(* IEC 61131-3 sources: daoli-st-library/DL_Device (part 24) *)

(* ---- FB_DL_HumidifierWaterQual.st ---- *)
(*
  FB_DL_HumidifierWaterQual  —  加湿器水质电导率监视与排水联锁 / Humidifier water conductivity monitoring with drain interlock
  分类 Category : DL_Device
  码位 Code     : 16#03_2_04
  版本 Version  : 1.0.0
  溯源 Source   : 道莅自研 clean-room（电导率标定与排水联锁为通用水处理工程语义）
  功能 Function : 1) 电导率经标定换算（斜率/偏置）后按门限分级，超标触发排水周期；
                  2) 排水阀与补水阀互斥，同拍双开即判冲突并双双回安全位（关阀）；
                  3) 电导门限带迟滞防抖，越限解除有可到达路径；标定斜率非法（0/负）即拒算并置码。
  边界 Boundary : ① 标定参数非法（斜率 0 或负）拒算并置码；
                  ② 排水联锁与补水阀互斥（同拍双开判冲突回安全位）；
                  ③ 电导门限带迟滞防抖，越限解除有可到达路径；
                  ④ 输出三行同向：电导值 → 分级 → 排水阀。
  依赖 Depends  : FC_DL_LimitClassify（电导分级，每拍无条件调用）、FB_DL_TimeWindowCheck（排水维护时间窗，每拍无条件调用）

  码表 Error codes（本件子码步进 16#10，避让邻件码位）:
    16#0002_0304 故障级：电导率标定参数非法（斜率 <= 0 或非有限），拒算
    16#0002_0314 故障级：排水阀与补水阀同拍双开（互斥冲突），双双回安全位
    16#0002_0324 信息级：电导率越限已启动排水（不置 bError）
*)

TYPE E_DL_HwqPhase :
(
    eIdle    := 0,   // 空闲 / Idle
    eMonitor := 10,  // 电导监视 / Conductivity monitoring
    eDrain   := 20,  // 排水周期进行 / Drain cycle running
    eHold    := 30,  // 拒算保持 / Rejected, held
    eFault   := 90   // 故障锁定 / Fault locked
);
END_TYPE

FUNCTION_BLOCK FB_DL_HumidifierWaterQual
VAR_INPUT
    bEnable      : BOOL;                          // 总使能，FALSE 关阀回空闲 / Master enable
    bReset       : BOOL;                          // 复位，上升沿清故障与冲突锁存 / Reset
    fCondRawUScm : REAL;                          // 电导率原始值 [uS/cm]，域 0~2000 / Raw conductivity [uS/cm]
    fCalSlope    : REAL := 1.0;                   // 电导标定斜率 [uS/cm per 原始计数]，域 > 0 / Calibration slope
    fCalOffset   : REAL := 0.0;                   // 电导标定偏置 [uS/cm] / Calibration offset [uS/cm]
    fCondWarnUScm: REAL := 300.0;                 // 电导警告门限 [uS/cm]，域 > 0 / Conductivity warning limit
    fCondTripUScm: REAL := 600.0;                 // 电导排水门限 [uS/cm]，须 > 警告门限 / Drain trigger limit
    fCondHystUScm: REAL := 20.0;                  // 电导迟滞 [uS/cm]，域 >= 0 / Conductivity hysteresis
    tDrainTime   : TIME := T#30S;                 // 单次排水时长 [ms]，域 > 0 / Drain duration [ms]
    tDrainPeriod : TIME := T#10M;                 // 排水周期 [ms]，域 > 0 / Drain period [ms]
    uHourNow     : USINT := 0;                    // 当前时刻-时 [h]（注入，禁读 CPU 钟）/ Injected hour [h]
    uMinNow      : USINT := 0;                    // 当前时刻-分 [min]（注入）/ Injected minute [min]
    fEps         : REAL := 1.0E-6;                // 浮点判零容差 [1] / Floating zero tolerance
END_VAR
VAR_OUTPUT
    fCondUScm    : REAL;                          // 标定后电导率 [uS/cm] / Calibrated conductivity [uS/cm]
    bDrainValve  : BOOL;                          // 排水阀 [开关] / Drain valve
    bFillValve   : BOOL;                          // 补水阀 [开关] / Make-up fill valve
    bCondWarn    : BOOL;                          // 电导警告（保持型）/ Conductivity warning, held
    bInDrainWin  : BOOL;                          // 处于维护排水时间窗 / Inside maintenance drain window
    bValveConflict : BOOL;                        // 阀门互斥冲突标志 / Valve exclusion conflict flag
    bError       : BOOL;                          // 故障标志，与故障级码配对 / Fault flag paired with fault codes
    uErrorId     : UDINT;                         // 事件码，0 = 无事件 / Event code, 0 = none
    eStateOut    : E_DL_HwqPhase;                 // 状态机当前态，段尾单点映射 / Phase mapped at tail
END_VAR
VAR
    _eState      : E_DL_HwqPhase := E_DL_HwqPhase.eIdle;  // 内部状态 / Internal state
    rtrReset     : R_TRIG;                        // 复位沿 / Reset edge
    tonDrain     : TON;                           // 排水时长计时（自复位）/ Drain duration timer
    tonPeriod    : TON;                           // 排水周期节拍（自复位）/ Drain period tick
    fbWindow     : FB_DL_TimeWindowCheck;         // 排水维护时间窗实例（无条件调用）/ Drain time window
    bCalOk       : BOOL;                          // 标定参数合法 / Calibration valid
    bCfgOk       : BOOL;                          // 组态合法 / Configuration valid
    eBand        : E_DL_LimitBand;                // 电导分级结果 / Conductivity band
    aDayEn       : ARRAY[1..7] OF BOOL;           // 星期使能表（周一~周日）/ Weekday enable table
    nDay         : INT;                           // 星期填充下标 / Weekday fill index
    fCondCal     : REAL;                          // 标定后电导率暂存 [uS/cm] / Calibrated conductivity buffer
    bCondHigh    : BOOL;                          // 越排水门限标志 / Above drain threshold
    bDrainCmd    : BOOL;                          // 排水指令暂存 / Drain command buffer
    bFillCmd     : BOOL;                          // 补水指令暂存 / Fill command buffer
    uFault       : UDINT;                         // 锁存故障码 / Latched fault code
    uInfo        : UDINT;                         // 信息级码 / Information code
END_VAR
VAR CONSTANT
    DL_HWQ_CMAX  : REAL := 2000.0;                // 电导物理域上限 [uS/cm] / Conductivity domain high
END_VAR

(* === 段 0 · 实例刷新（无条件周期调用，自复位节拍）=== *)
rtrReset(CLK := bReset);                          // 每拍刷新复位沿
tonDrain(IN := (_eState = E_DL_HwqPhase.eDrain) AND (NOT tonDrain.Q), PT := tDrainTime);   // 自复位
tonPeriod(IN := NOT tonPeriod.Q, PT := tDrainPeriod);                                      // 周期心跳自复位
FOR nDay := 1 TO 7 DO
    aDayEn[nDay] := TRUE;                         // 维护排水窗与星期无关：全周使能
END_FOR
fbWindow(uHourNow := uHourNow,                    // 注入当前时
         uMinNow := uMinNow,                      // 注入当前分
         bEnableDay := TRUE,                      // 日窗使能
         aWeekdayEnable := aDayEn,                // 周一到周日全开（本地数组填充）
         uWeekdayNow := 1,                        // 星期注入（维护窗与星期无关）
         uHourOn := 0,                            // 窗开 00:00
         uMinOn := 0,                             // 窗开 0 分
         uHourOff := 23,                          // 窗关 23:00
         uMinOff := 59,                           // 窗关 59 分
         bReset := rtrReset.Q);                   // 复位沿清信息码
bInDrainWin := fbWindow.bInWindow;                // 时间窗输出

(* === 段 1 · 标定与组态闸 === *)
bCalOk := (fCalSlope > fEps) AND (fCalSlope = fCalSlope) AND (fCalOffset = fCalOffset);   // 斜率正域 + NaN 自反
bCfgOk := (fCondWarnUScm > fEps) AND (fCondTripUScm > fCondWarnUScm)
          AND (fCondHystUScm >= 0.0) AND (tDrainTime > T#0MS) AND (tDrainPeriod > T#0MS)
          AND (fCondWarnUScm = fCondWarnUScm) AND (fCondTripUScm = fCondTripUScm);   // 含 NaN 自反
IF NOT bCalOk THEN
    uFault := 16#0002_0304;                       // 故障级：标定参数非法，拒算
END_IF
IF NOT bCfgOk THEN
    uFault := 16#0002_0304;                       // 故障级：组态非法同码段（防无码可查）
END_IF
IF rtrReset.Q AND bCalOk AND bCfgOk THEN
    uFault := 16#0000;                            // 复位沿清锁存（复位路径可达）
    bValveConflict := FALSE;                      // 冲突标志同步复位
    bCondWarn := FALSE;                           // 警告标志同步复位
END_IF
uInfo := 16#0000;                                 // 信息码每拍清零
IF bCalOk AND (fCondRawUScm = fCondRawUScm) AND (fCondRawUScm >= 0.0)
   AND (fCondRawUScm <= DL_HWQ_CMAX) THEN
    fCondCal := fCondRawUScm * fCalSlope + fCalOffset;   // 标定换算
    IF fCondCal < 0.0 THEN
        fCondCal := 0.0;                          // 负电导截零（物理不可达）
    END_IF
    fCondUScm := fCondCal;                        // 电导值输出
ELSE
    fCondCal := 0.0;                              // 拒算：不出数值
END_IF

(* === 段 2 · 电导分级（函数每拍无条件调用）=== *)
eBand := FC_DL_LimitClassify(fVal := fCondCal,
                             fLowLimit := -1.0,               // 低低限：本件不使用（负值域）
                             fLowWarn := -0.5,                // 低警告限：本件不使用
                             fUpWarn := fCondWarnUScm,        // 高警告限
                             fUpLimit := fCondTripUScm);      // 高排水限
bCondHigh := (eBand = E_DL_LimitBand.eUpTripped);  // 到达排水级
IF eBand = E_DL_LimitBand.eUpWarn THEN
    bCondWarn := TRUE;                             // 警告级：置警告
END_IF

(* === 段 3 · 主状态机（ENUM + CASE，含 ELSE 兜底）=== *)
CASE _eState OF
E_DL_HwqPhase.eIdle :
    bDrainCmd := FALSE;                            // 空闲不排水
    bFillCmd := FALSE;                             // 空闲不补水
    IF (uFault <> 16#0000) AND (uFault <> 16#0002_0314) THEN
        _eState := E_DL_HwqPhase.eFault;           // 故障优先
    ELSIF bEnable AND (NOT bCalOk) THEN
        _eState := E_DL_HwqPhase.eHold;            // 标定非法：拒算保持
    ELSIF bEnable THEN
        _eState := E_DL_HwqPhase.eMonitor;         // 进入监视相
    END_IF

E_DL_HwqPhase.eMonitor :
    bFillCmd := NOT bDrainCmd;                     // 补水默认开（与排水互斥）
    IF bCondHigh THEN
        bCondWarn := TRUE;                         // 置位型：电导警告
        uInfo := 16#0002_0324;                     // 信息级：越限启动排水
        _eState := E_DL_HwqPhase.eDrain;           // 转排水相
    ELSIF (eBand = E_DL_LimitBand.eNormal) AND (fCondCal < (fCondWarnUScm - fCondHystUScm)) THEN
        bCondWarn := FALSE;                        // 迟滞带下方：解除警告（可到达的解除路径）
    END_IF
    IF (NOT bEnable) OR (NOT bCalOk) THEN
        _eState := E_DL_HwqPhase.eIdle;            // 失能/标定失效回空闲
    END_IF

E_DL_HwqPhase.eDrain :
    bDrainCmd := TRUE;                             // 排水阀开（驱动方向）
    bFillCmd := FALSE;                             // 补水阀关（互斥）
    IF tonDrain.Q THEN
        bDrainCmd := FALSE;                        // 排水时长到：关阀（本拍行为）
        IF bCondHigh THEN
            IF tonPeriod.Q THEN
                bFillCmd := TRUE;                  // 周期未到且仍超标：等待下一周期再排
            END_IF
            _eState := E_DL_HwqPhase.eMonitor;     // 回监视相，等下一周期
        ELSE
            _eState := E_DL_HwqPhase.eMonitor;     // 达标：回监视相
        END_IF
    END_IF

E_DL_HwqPhase.eHold :
    bDrainCmd := FALSE;                            // 拒算态关排水
    bFillCmd := FALSE;                             // 拒算态关补水
    IF bCalOk THEN
        _eState := E_DL_HwqPhase.eMonitor;         // 标定恢复：解除拒算（可到达的解除路径）
    END_IF

E_DL_HwqPhase.eFault :
    bDrainCmd := FALSE;                            // 故障态排水阀关（安全侧）
    bFillCmd := FALSE;                             // 故障态补水阀关
    IF uFault = 16#0000 THEN
        _eState := E_DL_HwqPhase.eIdle;            // 解锁回空闲
    END_IF

ELSE
    _eState := E_DL_HwqPhase.eFault;               // 非法状态拦截
    uFault := 16#0002_0304;                        // 故障级：相 ID 越界
    bDrainCmd := FALSE;                            // 安全侧关阀
    bFillCmd := FALSE;                             // 安全侧关阀
END_CASE

(* === 段 4 · 阀门互斥仲裁（同拍双开判冲突，双双回安全位）=== *)
IF bDrainCmd AND bFillCmd THEN
    bDrainCmd := FALSE;                            // 冲突：排水阀回安全位
    bFillCmd := FALSE;                             // 冲突：补水阀回安全位
    bValveConflict := TRUE;                        // 冲突标志置位
    uFault := 16#0002_0314;                        // 故障级：互斥冲突
ELSE
    bValveConflict := FALSE;                       // 无冲突：标志清零（非置位型）
END_IF
IF rtrReset.Q AND bValveConflict THEN
    uFault := 16#0000;                             // 冲突经复位解除（复位路径可达）
    bValveConflict := FALSE;                       // 标志同步清零
END_IF
IF NOT bEnable THEN
    bDrainCmd := FALSE;                            // 失能最高优先：排水关
    bFillCmd := FALSE;                             // 失能最高优先：补水关
END_IF

(* === 段 5 · 输出映射（三行同向：电导值 → 分级 → 排水阀）=== *)
bDrainValve := bDrainCmd;                          // 排水阀输出
bFillValve := bFillCmd;                            // 补水阀输出
bError := (uFault <> 16#0000);                     // 故障标志仅由故障级码置位（R45 配对）
IF bError THEN
    uErrorId := uFault;                            // 故障级优先上报
ELSE
    uErrorId := uInfo;                             // 否则上报信息级码
END_IF
eStateOut := _eState;                              // 输出枚举段尾单点映射（N2 规则）
END_FUNCTION_BLOCK

(* ---- FB_DL_HydraulicAccumPreChg.st ---- *)
(*
  ==================================================================
  组件名 Component  : FB_DL_HydraulicAccumPreChg
  分类   Category   : DL_Device
  复杂度 Complexity  : cx3
  版本   Version    : 1.0.1
  功能   Purpose    : 液压蓄能器氮气预充压力监视。把实测气囊压力按理想气体等温
                      折算到参考温度 20 摄氏度（pCorr = pGas · T0K / TK），再对额定
                      预充压力求偏差百分比；欠充 / 过充双态判据带迟滞防抖；油口
                      压力显著高于气囊侧判气囊失效疑点（eBladderSuspect）；传感器
                      非有限或压力 / 温度物理域越界判 eSensorBad。
  来源   Source     : t2-2-lbp
  溯源   Origin     : IEC 61131-3 标准语义的道莅防御性实现；理想气体等温折算与
                      蓄能器预充校验为公开热力学与液压语义，clean-room 自研实现，
                      未复制任何闭源代码行。
  平台   Platform   : 纯 IEC 61131-3（LREAL 运算，无私有库、无定时器实例）
  作者   Author     : 道莅代码库 · PLC 编程专家（R56）
  ------------------------------------------------------------------
  边界 Boundary     :
                      一 本件只做预充状态判级，不做充放气控制、不做泄放（属主边界）；
                      二 判据方向性（R146）：欠充与过充为同量纲双向异常，分派独立
                         成因成员（R190 归因唯一），互不合并；
                      三 迟滞口径：进入判据用全带宽，退出判据带宽收窄 fHystBar，
                         防边界抖动反复置清；
                      四 成因锁存解除路径 = bReset 上升沿（唯一路径，头注释声明，R188）；
                      五 无全局变量、无外部变量声明、无物理地址寻址。
  输出契约 Output contract:
                      fDevPct 为温度修正后偏差百分比（正 = 高于额定，负 = 低于额定）；
                      eFault 为锁存回放；bError 与故障级成因配对（R45）；
                      ePhaseBad 为非法相位兜底专用成员（R128）。
  修订记录 Revision  :
    2026-11-20  v1.0.0  R56 首版（批 2 · 序号 10）
    2026-11-21  v1.0.1  R57 返修：段 3 域闸补温度上界 150.0 摄氏度判 eSensorBad（阈值提为常量并注单位）
  ==================================================================
*)

TYPE E_DL_HapPhase :
(
    eIdle  := 0,  // 未使能：判级停摆 / disabled, the grading is idle
    eRun   := 10, // 运行：逐拍判级 / running, graded every scan
    eFault := 90  // 故障：成因锁存 / fault, the cause is latched
);
END_TYPE

TYPE E_DL_HapFault :
(
    eNone          := 0, // 无成因 / no cause
    eUnderCharge   := 1, // 预充不足（故障级，与 bError 配对）/ the precharge is under, fault grade paired with bError
    eOverCharge    := 2, // 预充过量（故障级，与 bError 配对）/ the precharge is over, fault grade paired with bError
    eBladderSuspect:= 3, // 油口压力显著高于气囊侧，气囊失效疑点（故障级，与 bError 配对）/ the oil side clearly exceeds the gas side, a bladder suspect, fault grade paired with bError
    eSensorBad     := 4, // 传感器非有限或物理域越界（故障级，与 bError 配对）/ a sensor is non finite or out of the physical domain, fault grade paired with bError
    ePhaseBad      := 5  // 非法相位兜底（故障级，与 bError 配对）/ illegal phase fallback, fault grade paired with bError
);
END_TYPE

FUNCTION_BLOCK FB_DL_HydraulicAccumPreChg
VAR_INPUT
    bEnable   : BOOL := TRUE;   // 使能，失能时判级停摆 [-] / enable, the grading stops when disabled
    bReset    : BOOL := FALSE;  // 复位上升沿清全部成因锁存 [-] / reset rising edge clears every cause latch
    pGas      : LREAL := 90.0;  // 气囊压力实测 [巴] / measured gas side pressure [bar]
    pOil      : LREAL := 0.0;   // 油口压力实测 [巴] / measured oil port pressure [bar]
    fTempC    : LREAL := 20.0;  // 气体温度实测 [摄氏度] / measured gas temperature [degree celsius]
    pNom      : LREAL := 90.0;  // 额定预充压力 [巴]，域 大于零 / rated precharge pressure [bar], domain above zero
    fUnderBar : LREAL := 9.0;   // 欠充判据带宽（低于额定的绝对量）[巴] / undercharge band below the rating [bar]
    fOverBar  : LREAL := 9.0;   // 过充判据带宽（高于额定的绝对量）[巴] / overcharge band above the rating [bar]
    fHystBar  : LREAL := 1.0;   // 迟滞带宽 [巴]，域 0..判据带宽 / hysteresis band [bar], inside the criterion band
    fBladMarg : LREAL := 20.0;  // 气囊疑点裕度（油口超出气囊侧百分比）[百分比] / bladder suspect margin over the gas side [percent]
END_VAR
VAR_OUTPUT
    fDevPct : LREAL := 0.0;  // 温度修正后预充偏差百分比 [百分比] / the corrected precharge deviation [percent]
    ePhase  : E_DL_HapPhase := E_DL_HapPhase.eIdle; // 相位出口 [枚举] / phase outlet [enum]
    eFault  : E_DL_HapFault := E_DL_HapFault.eNone; // 成因出口，锁存回放 [枚举] / cause outlet replayed from the latch [enum]
    bError  : BOOL := FALSE; // 故障锁存标志 [-] / fault latch flag
END_VAR
VAR
    rtReset  : R_TRIG; // 复位沿检测，段 0 无条件刷新 / reset edge, refreshed unconditionally in segment zero
    _ePhase  : E_DL_HapPhase := E_DL_HapPhase.eIdle; // 内部相位，CASE 唯一写入目标 / internal phase, the only CASE write target
    _eFaulC  : E_DL_HapFault := E_DL_HapFault.eNone; // 故障级成因，锁存至复位沿 / fault cause, latched until the reset edge
    _bFault  : BOOL := FALSE; // 故障锁存位 [-] / fault latch bit
    _bInit   : BOOL := FALSE; // 首扫初始化完成标志（R310）/ first scan initialisation flag
    _bInOk   : BOOL := FALSE; // 三个实数输入全部有限 [-] / all three real inputs are finite
    _bCfgOk  : BOOL := FALSE; // 组态参数域内 [-] / the configuration is inside the domain
    _fTK     : LREAL := 0.0;  // 气体绝对温度 [开尔文] / the absolute gas temperature [kelvin]
    _fPCorr  : LREAL := 0.0;  // 折算到参考温度的气囊压力 [巴] / the gas pressure corrected to the reference temperature [bar]
    _fDev    : LREAL := 0.0;  // 偏差绝对量 [巴] / the deviation magnitude [bar]
    _bUnder  : BOOL := FALSE; // 欠充迟滞锁存 [-] / the undercharge hysteresis latch
    _bOver   : BOOL := FALSE; // 过充迟滞锁存 [-] / the overcharge hysteresis latch
    _bBlad   : BOOL := FALSE; // 气囊疑点迟滞锁存 [-] / the bladder suspect hysteresis latch
    _bBad    : BOOL := FALSE; // 传感器无效锁存 [-] / the sensor bad latch
END_VAR
VAR CONSTANT
    DL_HAP_TEMP_HI : LREAL := 150.0; // 温度上界 [摄氏度]，超界判传感器无效（v1.0.1 返修）/ the temperature ceiling [degree celsius], beyond it the sensor is judged bad (v1.0.1 fix)
END_VAR

// 段 0｜沿检测无条件周期刷新（禁入分支）/ segment 0, unconditional refresh of the edge detector
rtReset(CLK := bReset); // 复位沿无条件刷新 / unconditional refresh of the reset edge

// 段 1｜首扫初始化（R310）/ segment 1, first scan initialisation
IF NOT _bInit THEN // 首扫一拍 / the very first scan
    _bInit := TRUE; // 置首扫完成标志 / raise the first scan flag
    _ePhase := E_DL_HapPhase.eRun; // 相位从运行起步（使能默认真）/ the phase starts in run
    _eFaulC := E_DL_HapFault.eNone; // 故障级成因清零 / clear the fault cause
    _bFault := FALSE; // 故障锁存清零 / clear the fault latch
END_IF

// 段 2｜复位沿作用域：清全部迟滞与锁存 / 迁相位（两项逐项声明）/ segment 2, reset edge scope declared item by item
IF rtReset.Q THEN // 复位沿 / the reset edge
    _bFault := FALSE; // 作用域一：清故障锁存 / scope one, clear the fault latch
    _eFaulC := E_DL_HapFault.eNone; // 作用域一：清故障级成因 / scope one, clear the fault cause
    _bUnder := FALSE; // 作用域一：清欠充迟滞 / scope one, clear the undercharge latch
    _bOver := FALSE; // 作用域一：清过充迟滞 / scope one, clear the overcharge latch
    _bBlad := FALSE; // 作用域一：清气囊疑点迟滞 / scope one, clear the bladder latch
    _bBad := FALSE; // 作用域一：清传感器无效锁存 / scope one, clear the sensor bad latch
    _ePhase := E_DL_HapPhase.eRun; // 作用域二：迁回运行相 / scope two, migrate back to run
END_IF

// 段 3｜组态与输入域闸（R151 全覆盖）/ segment 3, the configuration and input domain gates
_bInOk := (pGas = pGas) AND ((pGas - pGas) = (pGas - pGas)) AND (pOil = pOil) AND ((pOil - pOil) = (pOil - pOil)) AND (fTempC = fTempC) AND ((fTempC - fTempC) = (fTempC - fTempC)); // 三输入有限性 / finiteness of the three inputs
_bCfgOk := (pNom > 0.0) AND (pNom = pNom) AND (fUnderBar >= 0.0) AND (fUnderBar = fUnderBar) AND (fOverBar >= 0.0) AND (fOverBar = fOverBar) AND (fHystBar >= 0.0) AND (fHystBar <= fUnderBar) AND (fHystBar <= fOverBar) AND (fBladMarg > 0.0) AND (fBladMarg = fBladMarg); // 组态参数域判定 / the configuration domain verdict
IF (NOT _bInOk) OR (pGas < 0.0) OR (pOil < 0.0) OR (fTempC < -270.0) OR (fTempC > DL_HAP_TEMP_HI) OR (NOT _bCfgOk) THEN // 输入非有限、物理域越界（含 v1.0.1 温度上界）或组态非法 / a non finite input, a physical domain violation (with the v1.0.1 temperature ceiling) or an illegal configuration
    IF NOT _bBad THEN // 未锁存才置（防同拍抹除）/ set only while unlatched
        _bBad := TRUE; // 置传感器无效锁存 / raise the sensor bad latch
    END_IF
END_IF

// 段 4｜相位机：ENUM + CASE，含 ELSE 非法相位兜底（R128）/ segment 4, the phase machine with an ELSE fallback
CASE _ePhase OF
E_DL_HapPhase.eIdle: // 未使能相 / the disabled phase
    IF bEnable AND (NOT _bFault) THEN // 使能且无故障 / enabled and unfaulted
        _ePhase := E_DL_HapPhase.eRun; // 迁运行相 / migrate to run
    END_IF

E_DL_HapPhase.eRun: // 运行相：逐拍判级 / the run phase, graded every scan
    IF NOT bEnable THEN // 失能 / disabled
        _ePhase := E_DL_HapPhase.eIdle; // 迁未使能相 / migrate to idle
    ELSIF _bBad THEN // 传感器无效锁存优先 / the sensor bad latch takes priority
        _bFault := TRUE; // 置故障锁存 / raise the fault latch
        _eFaulC := E_DL_HapFault.eSensorBad; // 故障级成因（R45 配对 bError）/ the fault cause paired with bError
        _ePhase := E_DL_HapPhase.eFault; // 迁故障相 / migrate to the fault phase
    ELSE // 正常判级 / the normal grading
        _fTK := fTempC + 273.15; // 摄氏度转开尔文 / celsius to kelvin
        IF _fTK < 1.0 THEN // 绝对温度趋零防御（等温折算除子域闸）/ the absolute temperature guard for the divisor
            _fTK := 1.0; // 钳到下限 / clamp to the floor
        END_IF
        _fPCorr := pGas * (293.15 / _fTK); // 等温折算到 20 摄氏度参考（除子为绝对温度已证超阈）/ the isothermal correction to the twenty degree reference
        IF pNom > 0.0 THEN // 额定压力已证大于零（组态闸）/ the rating is proven positive by the gate
            fDevPct := (_fPCorr - pNom) / pNom * 100.0; // 偏差百分比 / the deviation percentage
        ELSE // 组态非法兜底（防御性保留）/ the illegal configuration fallback
            fDevPct := 0.0; // 偏差记零 / the deviation is zeroed
        END_IF
        _fDev := _fPCorr - pNom; // 偏差绝对量（带符号）/ the signed deviation
        IF _fDev < -fUnderBar THEN // 欠充进入判据 / the undercharge entry criterion
            _bUnder := TRUE; // 置欠充迟滞锁存 / raise the undercharge latch
        ELSIF _fDev > -fUnderBar + fHystBar THEN // 欠充退出判据（迟滞收窄）/ the undercharge exit criterion with the narrowed band
            _bUnder := FALSE; // 清欠充迟滞 / clear the undercharge latch
        END_IF
        IF _fDev > fOverBar THEN // 过充进入判据 / the overcharge entry criterion
            _bOver := TRUE; // 置过充迟滞锁存 / raise the overcharge latch
        ELSIF _fDev < fOverBar - fHystBar THEN // 过充退出判据（迟滞收窄）/ the overcharge exit criterion with the narrowed band
            _bOver := FALSE; // 清过充迟滞 / clear the overcharge latch
        END_IF
        IF pOil > _fPCorr * (1.0 + fBladMarg / 100.0) THEN // 油口显著高于气囊侧 / the oil side clearly exceeds the gas side
            _bBlad := TRUE; // 置气囊疑点迟滞锁存 / raise the bladder latch
        ELSIF pOil < _fPCorr * (1.0 + fBladMarg / 200.0) THEN // 气囊疑点退出判据（半带迟滞）/ the bladder exit criterion with a half band
            _bBlad := FALSE; // 清气囊疑点迟滞 / clear the bladder latch
        END_IF
        IF _bBlad THEN // 气囊疑点优先级最高（结构性失效）/ the bladder suspect has the highest priority, a structural failure
            _bFault := TRUE; // 置故障锁存 / raise the fault latch
            _eFaulC := E_DL_HapFault.eBladderSuspect; // 故障级成因（R45 配对 bError）/ the fault cause paired with bError
            _ePhase := E_DL_HapPhase.eFault; // 迁故障相 / migrate to the fault phase
        ELSIF _bOver THEN // 过充次优先 / the overcharge takes the next priority
            _bFault := TRUE; // 置故障锁存 / raise the fault latch
            _eFaulC := E_DL_HapFault.eOverCharge; // 故障级成因（R45 配对 bError）/ the fault cause paired with bError
            _ePhase := E_DL_HapPhase.eFault; // 迁故障相 / migrate to the fault phase
        ELSIF _bUnder THEN // 欠充再次优先 / the undercharge follows
            _bFault := TRUE; // 置故障锁存 / raise the fault latch
            _eFaulC := E_DL_HapFault.eUnderCharge; // 故障级成因（R45 配对 bError）/ the fault cause paired with bError
            _ePhase := E_DL_HapPhase.eFault; // 迁故障相 / migrate to the fault phase
        END_IF
    END_IF

E_DL_HapPhase.eFault: // 故障相：成因锁存，等待复位沿；偏差出口冻结保持末值（R191 显式声明）/ the fault phase, the cause is latched, the deviation outlet holds frozen

ELSE // 非法相位兜底（R128）/ the illegal phase fallback
    _bFault := TRUE; // 置故障锁存 / raise the fault latch
    _eFaulC := E_DL_HapFault.ePhaseBad; // 故障级成因（R45 配对 bError）/ the fault cause paired with bError
    _ePhase := E_DL_HapPhase.eFault; // 迁故障相 / migrate to the fault phase
END_CASE

// 段 5｜统一出口 / segment 5, the unified outlet
IF _bFault THEN // 故障锁存优先 / the fault latch takes priority
    eFault := _eFaulC; // 故障级成因锁存回放（不按当下输入重推断，R152）/ the fault cause replayed from the latch
ELSE
    eFault := E_DL_HapFault.eNone; // 无锁存即无成因 / no latch, no cause
END_IF
ePhase := _ePhase; // 相位出口单点映射 / single point phase outlet mapping
bError := _bFault; // 故障标志与锁存位同源 / the fault flag shares the latch source
END_FUNCTION_BLOCK

(* ---- FB_DL_HydroPressRampSeq.st ---- *)
(*
  ============================================================
  组件名 : FB_DL_HydroPressRampSeq
  分类   : DL_Device
  功能   : 液压建压斜坡顺序控制，建压升压保压泄压按斜率给定并含超时保护
  开源溯源 : internal-design（本轮无外部代码逐行引用）
             参考语义 : 无外部参考
  复杂度 : C2
  版本   : 1.0.0
  ============================================================
  配比约束 : tonRamp 与 tonHold 共用 tHoldTimeout 作为监视窗（升压窗与保压窗各一实例，
             两者互不累计）；tReleaseTimeout 单独覆盖泄压相。默认值须全部大于零。
  降级语义 : 实测压力非有限时冻结斜坡并保持上一有限设定输出，bPressOk 置假，不置故障码。
  故障码   : 1 保压超时 / 2 升压超时 / 3 泄压超时。码 3 不可由 1 与 2 观测——1 与 2 只在
             升压相与保压相置位，泄压相进入故障时码必为 0，故单开 3 以区分成因。
             复位唯一路径：bBuildCmd 或 bReleaseCmd 上升沿。
  ============================================================
*)

TYPE E_DL_HydroRampState :
(
    eIdle     := 0, // 待机，设定保持在零 idle with the set point at zero
    eRampUp   := 1, // 升压相，按斜率逼近目标 pressure ramp up towards the target
    eHold     := 2, // 保压相，设定保持目标 pressure hold at the target
    eRampDown := 3, // 泄压相，按斜率降到零 pressure ramp down to zero
    eFault    := 4  // 故障锁存相 latched fault phase
);
END_TYPE

FUNCTION_BLOCK FB_DL_HydroPressRampSeq
VAR_INPUT
    bBuildCmd      : BOOL; // 建压命令 pressure build command
    bReleaseCmd    : BOOL; // 泄压命令 pressure release command
    rPressAct      : REAL; // 实测压力 [bar] actual pressure [bar]
    rPressTarget   : REAL; // 目标压力 [bar] target pressure [bar]
    rRampBarPerS   : REAL; // 升压斜率 [bar/s] ramp rate [bar per second]
    rHoldBand      : REAL; // 保压允差带 [bar] hold band [bar]
    tHoldTimeout   : TIME; // 保压与升压监视窗 [ms] hold and ramp watchdog window
    tReleaseTimeout: TIME; // 泄压监视窗 [ms] release watchdog window
END_VAR
VAR_OUTPUT
    rPressSp   : REAL; // 压力设定输出 [bar] pressure set point [bar]
    eState     : E_DL_HydroRampState; // 当前状态 current state
    bPressOk   : BOOL; // 保压到位标志 pressure reached flag
    nFaultCode : INT; // 故障码 0无 1保压超时 2升压超时 3泄压超时 [码] fault code [code]
END_VAR
VAR
    _eState  : E_DL_HydroRampState := E_DL_HydroRampState.eIdle; // 内部状态 internal state
    _rSp     : REAL := 0.0; // 斜坡积分设定量 [bar] ramped set point [bar]
    _nFault  : INT := 0; // 故障码锁存内部量 latched fault code
    _bFin    : BOOL := FALSE; // 实数输入有限性判定 finiteness verdict of the real inputs
    _rBand   : REAL := 0.0; // 钳位后的允差带 [bar] clamped hold band [bar]
    tonTick  : TON; // 一秒节拍计时 one second tick timer
    tonHold  : TON; // 保压超时计时 hold timeout timer
    tonRamp  : TON; // 升压超时计时 ramp timeout timer
    tonRelease : TON; // 泄压超时计时 release timeout timer
    rtBuild  : R_TRIG; // 建压命令上升沿 build command rising edge
    rtRelease: R_TRIG; // 泄压命令上升沿 release command rising edge
END_VAR

// 段 0｜定时器与沿实例无条件周期刷新 unconditional cyclic refresh of timers and edges
tonTick(IN := NOT tonTick.Q, PT := T#1S); // 一秒自复位节拍 one second self reset tick
tonHold(IN := (_eState = E_DL_HydroRampState.eHold) AND (_nFault = 0), PT := tHoldTimeout); // 保压超时 hold timeout
tonRamp(IN := (_eState = E_DL_HydroRampState.eRampUp) AND (_nFault = 0), PT := tHoldTimeout); // 升压超时 ramp timeout
tonRelease(IN := (_eState = E_DL_HydroRampState.eRampDown) AND (_nFault = 0), PT := tReleaseTimeout); // 泄压超时 release timeout
rtBuild(CLK := bBuildCmd); // 建压沿刷新 refresh the build edge
rtRelease(CLK := bReleaseCmd); // 泄压沿刷新 refresh the release edge
// 段 1｜出口预置与输入整形 preset the outputs and reshape the inputs
bPressOk := FALSE; // 到位标志每拍先假 the reached flag is false each scan first
_rBand := rHoldBand; // 取入参允差带 take the hold band input
IF _rBand < 0.0 THEN
    _rBand := ABS(_rBand); // 负允差带取幅值 a negative band becomes its magnitude
END_IF
_bFin := (rPressAct = rPressAct) AND (rPressTarget = rPressTarget) AND (rRampBarPerS = rRampBarPerS) AND (rHoldBand = rHoldBand); // 四输入自反判定 self comparison of the four inputs
IF NOT _bFin THEN
    rPressSp := _rSp; // 冻结斜坡并输出上一有限设定 freeze the ramp and emit the last finite set point
    eState := _eState; // 状态出口按锁存量 map the state
    nFaultCode := _nFault; // 故障码出口按锁存量 map the fault code
    RETURN; // 非有限测量不迁相，早退 the non finite reading changes no phase
END_IF
// 段 2｜主状态机 main state machine
CASE _eState OF
E_DL_HydroRampState.eIdle: // 待机相 idle phase
    _rSp := 0.0; // 待机设定归零 the set point returns to zero
    IF rtBuild.Q AND (NOT bReleaseCmd) AND (rPressTarget > 0.0) AND (rRampBarPerS > 0.0) THEN
        _eState := E_DL_HydroRampState.eRampUp; // 组态合法才迁升压相 migrate only when the configuration is legal
    END_IF
E_DL_HydroRampState.eRampUp: // 升压相 ramp up phase
    IF tonTick.Q THEN
        _rSp := LIMIT(0.0, _rSp + rRampBarPerS, rPressTarget); // 每满一秒按斜率推进 advance one ramp step per full second
    END_IF
    IF (rPressAct >= (rPressTarget - _rBand)) AND (ABS(_rSp - rPressTarget) < 1.0E-3) THEN
        _eState := E_DL_HydroRampState.eHold; // 设定到位且反馈入带则迁保压 both the set point and the feedback are in place
    ELSIF tonRamp.Q THEN
        _nFault := 2; // 升压超时故障码 ramp timeout fault code
        _eState := E_DL_HydroRampState.eFault; // 迁故障相 migrate to the fault phase
    END_IF
E_DL_HydroRampState.eHold: // 保压相 hold phase
    _rSp := rPressTarget; // 设定保持目标 the set point holds the target
    IF ABS(rPressAct - rPressTarget) <= _rBand THEN
        bPressOk := TRUE; // 反馈在允差带内 the feedback sits inside the band
    END_IF
    IF rtRelease.Q OR bReleaseCmd THEN
        _eState := E_DL_HydroRampState.eRampDown; // 泄压命令优先于超时 the release command outranks the timeout
    ELSIF tonHold.Q THEN
        _nFault := 1; // 保压超时故障码 hold timeout fault code
        _eState := E_DL_HydroRampState.eFault; // 迁故障相 migrate to the fault phase
    END_IF
E_DL_HydroRampState.eRampDown: // 泄压相 ramp down phase
    IF tonTick.Q THEN
        _rSp := LIMIT(0.0, _rSp - rRampBarPerS, rPressTarget); // 每满一秒按斜率回落 fall one ramp step per full second
    END_IF
    IF (rPressAct < 0.5) AND (_rSp < 1.0E-3) THEN
        _rSp := 0.0; // 设定归零 the set point lands at zero
        _eState := E_DL_HydroRampState.eIdle; // 回待机 return to idle
    ELSIF tonRelease.Q THEN
        _nFault := 3; // 泄压超时故障码 release timeout fault code
        _eState := E_DL_HydroRampState.eFault; // 迁故障相 migrate to the fault phase
    END_IF
E_DL_HydroRampState.eFault: // 故障锁存相 latched fault phase
    IF rtBuild.Q OR rtRelease.Q THEN
        _nFault := 0; // 复位清故障码 the reset edge clears the fault code
        _rSp := 0.0; // 复位设定归零 the reset edge clears the set point
        _eState := E_DL_HydroRampState.eIdle; // 复位回待机 the reset edge returns to idle
    END_IF
ELSE // 非法状态枚举兜底 the illegal state fallback
    _eState := E_DL_HydroRampState.eIdle; // 非法状态回落待机 an illegal state falls back to idle
END_CASE
// 段 3｜统一出口映射 the unified exit mapping
rPressSp := _rSp; // 设定出口 map the set point
eState := _eState; // 状态出口 map the state
nFaultCode := _nFault; // 故障码出口 map the fault code
END_FUNCTION_BLOCK

(* ---- FB_DL_InductionHardeningScanCtrl.st ---- *)
(*
  Component : FB_DL_InductionHardeningScanCtrl
  Category  : DL_Device
  Type      : FB
  Complexity: C2
  VERSION   : v1.0.0
  功能      : 感应淬火扫描时序控制：ENUM 七态状态机（Idle/Heat/Scan/Spray/Cool/Done/Fault），扫描功率随速度联动，喷淋延时后转冷却。
  开源溯源  : 道莅原创 clean-room 自研（无外部代码引用）｜License: MIT
  边界条件  : ① 扫描速度设定/参考速度/终点行程为除子或比例基，须 > 1e-9，否则拒启动并锁存故障码；
              ② 功率按速度比线性联动并钳位 0~100 %，速度越界不下发超限功率；
              ③ 故障锁存唯一解除路径 = bReset 上升沿；eDone 撤销 bStart 回 eIdle。
*)

TYPE E_DL_IhScanPhase :
(
    eIdle  := 0,    (* 空闲：等启动沿 / Idle waiting start edge *)
    eHeat  := 10,   (* 预热：定时加热 / Pre-heating by timer *)
    eScan  := 20,   (* 扫描：速度功率联动 / Scanning with speed-power link *)
    eSpray := 30,   (* 喷淋：延时后开喷 / Spray after delay *)
    eCool  := 40,   (* 冷却：驻留冷却 / Cooling dwell *)
    eDone  := 50,   (* 完成：结论驻留 / Done, result held *)
    eFault := 90    (* 故障：锁存待复位 / Fault latched *)
);
END_TYPE

FUNCTION_BLOCK FB_DL_InductionHardeningScanCtrl
VAR_INPUT
    bEnable         : BOOL;   (* 使能电平 [-] Enable level *)
    bReset          : BOOL;   (* 复位上升沿，清故障锁存 [-] Reset edge *)
    bStart          : BOOL;   (* 启动上升沿 [-] Start edge *)
    fScanPosMm      : REAL;   (* 感应器实际位置 [mm] Inductor actual position *)
    fScanEndMm      : REAL;   (* 扫描终点行程 [mm] Scan end stroke *)
    fScanSpeedSetMmS: REAL;   (* 扫描速度设定 [mm/s] Scan speed setpoint *)
    fSpeedRefMmS    : REAL;   (* 功率联动参考速度 [mm/s] Speed reference for power link *)
    fPowerSetPct    : REAL;   (* 额定功率设定 [%] Rated power setpoint *)
    tHeatDur        : TIME;   (* 预热驻留 [ms] Pre-heat dwell *)
    tSprayDelay     : TIME;   (* 喷淋开启延时 [ms] Spray on delay *)
    tCoolDur        : TIME;   (* 冷却驻留 [ms] Cooling dwell *)
END_VAR
VAR_OUTPUT
    bHeatOn      : BOOL;             (* 加热输出 [-] Heating output *)
    bScanRun     : BOOL;             (* 扫描运行输出 [-] Scan run output *)
    bSprayOn     : BOOL;             (* 喷淋输出 [-] Spray output *)
    fPowerOutPct : REAL;             (* 功率输出（速度联动后） [%] Power output after link *)
    fSpeedOutMmS : REAL;             (* 速度输出 [mm/s] Speed output *)
    ePhase       : E_DL_IhScanPhase; (* 相位出口，段尾单点映射 [-] Phase outlet *)
    bError       : BOOL;             (* 故障锁存标志 [-] Fault latch flag *)
    uErrId       : UDINT;            (* 事件码，0 = 无事件 [-] Event code *)
END_VAR
VAR
    rtReset   : R_TRIG;   (* 复位沿实例，每拍无条件刷新 / Reset edge *)
    rtStart   : R_TRIG;   (* 启动沿实例，每拍无条件刷新 / Start edge *)
    tonHeat   : TON;      (* 预热驻留计时（独立实例） / Pre-heat timer *)
    tonSpray  : TON;      (* 喷淋延时计时（独立实例） / Spray delay timer *)
    tonCool   : TON;      (* 冷却驻留计时（独立实例） / Cooling timer *)
    _ePhase   : E_DL_IhScanPhase := E_DL_IhScanPhase.eIdle;  (* 内部相位 / Internal phase *)
    _bFault   : BOOL;     (* 故障锁存位（锁存量） / Latched fault bit *)
    _uFault   : UDINT;    (* 故障码锁存（锁存量） / Latched fault code *)
    _bCfgBad  : BOOL;     (* 组态非法当拍量 [-] / Config illegal flag *)
    _bNonFin  : BOOL;     (* 输入非有限当拍量 [-] / Non-finite input flag *)
END_VAR
VAR CONSTANT
    DL_EPS     : REAL := 1.0E-9;   (* 除零判定容差 [无量纲] Divide-by-zero tolerance *)
    DL_PCT_MAX : REAL := 100.0;    (* 功率百分比上限 [%] Power percent upper bound *)
END_VAR

(* —— 段 0｜沿与定时器每拍无条件刷新（禁置于 IF/CASE 内，使能挂 IN 引脚） —— *)
rtReset(CLK := bReset);
rtStart(CLK := bStart);
tonHeat (IN := (_ePhase = E_DL_IhScanPhase.eHeat) AND (NOT _bFault), PT := tHeatDur);
tonSpray(IN := (_ePhase = E_DL_IhScanPhase.eSpray) AND (NOT _bFault), PT := tSprayDelay);
tonCool (IN := (_ePhase = E_DL_IhScanPhase.eCool) AND (NOT _bFault), PT := tCoolDur);

(* —— 段 1｜每拍量预清零（锁存量 _bFault/_uFault 不入清单） —— *)
uErrId := 16#0000_0000;
_bCfgBad := FALSE;
_bNonFin := FALSE;

(* —— 段 2｜复位沿：故障一次性清干净，相位回空闲，输出撤销 —— *)
IF rtReset.Q THEN
    _bFault := FALSE;
    _uFault := 16#0000_0000;
    _ePhase := E_DL_IhScanPhase.eIdle;
END_IF

(* —— 段 3｜组态闸：覆盖全部参与判据换算的引脚（速度/终点/功率/时长） —— *)
IF (fScanSpeedSetMmS <= DL_EPS) OR (fSpeedRefMmS <= DL_EPS)
   OR (fScanEndMm <= DL_EPS) OR (fPowerSetPct <= 0.0)
   OR (tHeatDur = T#0S) OR (tCoolDur = T#0S) THEN
    _bCfgBad := TRUE;
END_IF
IF (fScanPosMm <> fScanPosMm) OR ((fScanPosMm - fScanPosMm) <> 0.0)
   OR (fPowerSetPct <> fPowerSetPct) OR ((fPowerSetPct - fPowerSetPct) <> 0.0)
   OR (fScanSpeedSetMmS <> fScanSpeedSetMmS) OR ((fScanSpeedSetMmS - fScanSpeedSetMmS) <> 0.0)
   OR (fSpeedRefMmS <> fSpeedRefMmS) OR ((fSpeedRefMmS - fSpeedRefMmS) <> 0.0) THEN
    _bNonFin := TRUE;
END_IF

(* —— 段 4｜主状态机：七态全覆盖 + ELSE 兜底 —— *)
CASE _ePhase OF
E_DL_IhScanPhase.eIdle:
    bHeatOn := FALSE; bScanRun := FALSE; bSprayOn := FALSE;
    fPowerOutPct := 0.0; fSpeedOutMmS := 0.0;
    IF rtStart.Q AND bEnable AND (NOT _bFault) AND (NOT _bCfgBad) AND (NOT _bNonFin) THEN
        _ePhase := E_DL_IhScanPhase.eHeat;
    ELSIF rtStart.Q AND (_bFault OR _bCfgBad OR _bNonFin) THEN
        _bFault := TRUE;                 (* 带病启动拒绝 / Reject start with bad config *)
        _uFault := 16#0020_0001;         (* 故障级：组态非法 / Fault code bad config *)
        _ePhase := E_DL_IhScanPhase.eFault;
    END_IF

E_DL_IhScanPhase.eHeat:
    bHeatOn := TRUE; bScanRun := FALSE; bSprayOn := FALSE;
    fSpeedOutMmS := 0.0;
    IF _bNonFin THEN
        _bFault := TRUE; _uFault := 16#0020_0002;   (* 故障级：输入非有限 / Non-finite *)
        _ePhase := E_DL_IhScanPhase.eFault;
    ELSIF tonHeat.Q THEN
        _ePhase := E_DL_IhScanPhase.eScan;          (* 迁出条件 1：预热驻留完成 *)
    ELSIF NOT bEnable THEN
        _ePhase := E_DL_IhScanPhase.eIdle;          (* 迁出条件 2：使能撤销回安全态 *)
    END_IF

E_DL_IhScanPhase.eScan:
    bHeatOn := TRUE; bScanRun := TRUE; bSprayOn := FALSE;
    fSpeedOutMmS := fScanSpeedSetMmS;               (* 速度输出 = 设定值 [mm/s] *)
    (* 功率-速度联动：功率 = 额定功率 × 实际速度/参考速度，超限钳位 *)
    fPowerOutPct := fPowerSetPct * (fScanSpeedSetMmS / fSpeedRefMmS);
    IF fPowerOutPct > DL_PCT_MAX THEN
        fPowerOutPct := DL_PCT_MAX;                 (* 功率上限钳位 [%] / Power clamp *)
    ELSIF fPowerOutPct < 0.0 THEN
        fPowerOutPct := 0.0;                        (* 功率下限钳位 [%] / Power floor *)
    END_IF
    IF _bNonFin THEN
        _bFault := TRUE; _uFault := 16#0020_0002;   (* 故障级：输入非有限 / Non-finite *)
        _ePhase := E_DL_IhScanPhase.eFault;
    ELSIF fScanPosMm >= fScanEndMm THEN
        _ePhase := E_DL_IhScanPhase.eSpray;         (* 迁出条件 1：扫描终点达成 *)
    ELSIF fScanPosMm < 0.0 THEN
        _bFault := TRUE; _uFault := 16#0020_0003;   (* 故障级：位置反馈越界 / Position out of range *)
        _ePhase := E_DL_IhScanPhase.eFault;         (* 迁出条件 2（故障路） *)
    ELSIF NOT bEnable THEN
        _ePhase := E_DL_IhScanPhase.eIdle;          (* 迁出条件 3：使能撤销 *)
    END_IF

E_DL_IhScanPhase.eSpray:
    bHeatOn := FALSE; bScanRun := FALSE;
    fSpeedOutMmS := 0.0; fPowerOutPct := 0.0;
    bSprayOn := tonSpray.Q;                         (* 延时到才开喷 / Spray after delay *)
    IF tonSpray.Q THEN
        _ePhase := E_DL_IhScanPhase.eCool;          (* 迁出条件 1：喷淋延时完成 *)
    ELSIF NOT bEnable THEN
        _ePhase := E_DL_IhScanPhase.eIdle;          (* 迁出条件 2：使能撤销 *)
    END_IF

E_DL_IhScanPhase.eCool:
    bHeatOn := FALSE; bScanRun := FALSE; bSprayOn := TRUE;
    fSpeedOutMmS := 0.0; fPowerOutPct := 0.0;
    IF tonCool.Q THEN
        _ePhase := E_DL_IhScanPhase.eDone;          (* 迁出条件 1：冷却驻留完成 *)
    ELSIF NOT bEnable THEN
        _ePhase := E_DL_IhScanPhase.eIdle;          (* 迁出条件 2：使能撤销 *)
    END_IF

E_DL_IhScanPhase.eDone:
    bHeatOn := FALSE; bScanRun := FALSE; bSprayOn := FALSE;
    fSpeedOutMmS := 0.0; fPowerOutPct := 0.0;
    IF NOT bStart THEN
        _ePhase := E_DL_IhScanPhase.eIdle;          (* 启动指令撤销：回空闲 *)
    END_IF

E_DL_IhScanPhase.eFault:
    bHeatOn := FALSE; bScanRun := FALSE; bSprayOn := FALSE;
    fSpeedOutMmS := 0.0; fPowerOutPct := 0.0;       (* 故障相：全部输出走安全侧 *)

ELSE
    _bFault := TRUE;                                (* 兜底：非法相位锁存 *)
    _uFault := 16#0020_0009;
    _ePhase := E_DL_IhScanPhase.eFault;
END_CASE

(* —— 段 5｜相位与故障码出口单点映射 —— *)
ePhase := _ePhase;
bError := _bFault;
IF _bFault AND (_uFault <> 16#0000_0000) THEN
    uErrId := _uFault;                              (* 故障码锁存回放 / Latched fault replay *)
END_IF
END_FUNCTION_BLOCK

(* ---- FB_DL_InverterDeratingCtrl.st ---- *)
(*
  Component : FB_DL_InverterDeratingCtrl
  Category  : DL_Device
  Type      : FB
  Version   : 1.0.1
  CodeSeg   : 16#03_1_04
  Summary   : 逆变器温度/电压分段降额与功率限值：NE107 四态降额状态机，降额原因独立枚举上报。
              Inverter staged derating and power limit: NE107 four-state machine with a separate reason enum.
  溯源声明  : 仅借 NE107 分类与参数域，代码 clean-room（T2 借鉴件）
  边界安全  : 温度/电压非有限（NaN 自反 + Inf 上限）拦截，故障时强制转入停机安全相；
              阈值域闸（tDer1 < tDer2 < tStop，vMax > 0）防止整定倒置；
              状态机 ENUM + CASE 且 ELSE 回 Normal 降级路径；降额原因枚举与 _eState 分离不复用；
              CASE 内禁止给输出枚举赋值，段 3 统一映射；迟滞回差防阈值抖动。
  复用      : 无
*)

FUNCTION_BLOCK FB_DL_InverterDeratingCtrl
VAR_INPUT
    bRun     : BOOL;                    (* 使能，假则回 Normal 并封零 · Enable *)
    fTempC   : LREAL;                   (* 逆变器温度 [degC] · Inverter temperature *)
    fVoltV   : LREAL;                   (* 直流母线电压 [V] · DC link voltage *)
    fT1C     : LREAL := 70.0;           (* 一级降额温度阈 [degC] · Level 1 derating temp *)
    fT2C     : LREAL := 80.0;           (* 二级降额温度阈 [degC] · Level 2 derating temp *)
    fTStopC  : LREAL := 90.0;           (* 停机温度阈 [degC] · Stop temperature *)
    fVoltMaxV: LREAL := 850.0;          (* 电压降额阈 [V] · Voltage derating threshold *)
    fPowerNomKw: LREAL := 100.0;        (* 额定功率 [kW] · Nominal power *)
    fHysC    : LREAL := 3.0;            (* 温度回差 [degC] · Temperature hysteresis *)
    fEps     : LREAL := 1.0E-6;         (* 浮点判零容差 [实数域] · Floating zero tolerance *)
END_VAR
VAR_OUTPUT
    eMode      : (eMNormal := 0, eMDerat1 := 1, eMDerat2 := 2, eMStop := 3);    (* 相枚举输出 / Mode output enum *)
    eReason    : (eRsnNone := 0, eRsnOverTemp := 1, eRsnOverVolt := 2);         (* 降额原因枚举，与相枚举分离 / Reason enum, separate type *)
    fPowerLimKw: LREAL;                (* 功率限值输出 [kW] · Power limit output *)
    bDerating  : BOOL;                  (* 降额激活标志 · Derating active flag *)
    bError     : BOOL;                  (* 故障标志，与故障码配对 · Fault flag paired with codes *)
    uErrorId   : UDINT;                 (* 事件码 16#0000_0104，0 无事件 · Event code *)
END_VAR
VAR
    _eState : (eStNormal := 0, eStDer1 := 1, eStDer2 := 2, eStStop := 3);   (* 内部状态机，与输出枚举分离 / Internal state *)
    uCode   : WORD;     (* 码位暂存，每拍重算 [码] · Code staging *)
    bSigOk  : BOOL;     (* 输入有效标志 · Input validity flag *)
    bThrOk  : BOOL;     (* 阈值整定域标志 · Threshold tuning validity *)
    eRsn    : (eIRsnNone := 0, eIRsnOverTemp := 1, eIRsnOverVolt := 2);        (* 内部原因枚举，成员名加 I 前缀防重声明 / Internal reason enum, prefixed members *)
END_VAR
VAR CONSTANT
    DL_IDC_PCT1 : LREAL := 0.8;         (* 一级降额功率比 [比值] · Level 1 power ratio *)
    DL_IDC_PCT2 : LREAL := 0.5;         (* 二级降额功率比 [比值] · Level 2 power ratio *)
END_VAR

(* === 段 0 · 实例刷新 === *)
(* 无 TON/R_TRIG 实例：本件为阈值状态机；No timer instances, threshold state machine *)

(* === 段 1 · 输入校验与量程闸 === *)
uCode := 16#0000;                       // 每拍清码（可达清零基线）/ Clear codes each scan
bSigOk := (fTempC = fTempC) AND (fVoltV = fVoltV)                   // NaN 自反判据 / NaN reflexivity
          AND (ABS(fTempC) < 1.0E308) AND (ABS(fVoltV) < 1.0E308);  // Inf 上限判据 / Inf limit
bThrOk := (fT1C < fT2C) AND (fT2C < fTStopC) AND (fVoltMaxV > fEps) // 阈值倒置闸 / Threshold order gate
          AND (fPowerNomKw > fEps) AND (fHysC >= 0.0);              // 功率/回差域闸 / Power and hysteresis gates
IF NOT bSigOk OR NOT bThrOk THEN
    uCode := 16#0104;                   // 故障级：域外或整定倒置 / Fault: domain or tuning invalid
END_IF

(* === 段 2 · 主逻辑：NE107 四态降额状态机 === *)
IF NOT bRun THEN
    _eState := eStNormal;               (* 撤使能回 Normal，输出封零在段 3 / Back to normal on disable *)
    eRsn := eIRsnNone;
ELSIF NOT bSigOk THEN
    _eState := eStStop;                 (* 输入非有限强制停机安全相 / Non-finite forces the stop state *)
    eRsn := eIRsnOverTemp;
ELSIF NOT bThrOk THEN
    (* 整定倒置：保持当前相不迁移，段 3 报码 / Bad tuning: hold state, code in segment 3 *)
ELSE
    eRsn := eIRsnNone;                  (* 默认无原因 / Default no reason *)
    CASE _eState OF
        eStNormal:                      (* 正常相：越阈升相 / Normal: escalate on thresholds *)
            IF (fTempC > fTStopC) OR (fVoltV > fVoltMaxV) THEN
                _eState := eStDer2;     (* 拍 N 越阈，拍 N+1 生效二级降额 / To derating 2 *)
                IF fVoltV > fVoltMaxV THEN
                    eRsn := eIRsnOverVolt;  (* 过压触发须归因过压，不得归因过温 / Over-volt attribution *)
                ELSE
                    eRsn := eIRsnOverTemp;  (* 过温触发归因过温 / Over-temp attribution *)
                END_IF
            ELSIF fTempC > fT1C THEN
                _eState := eStDer1;     (* 拍 N+1 一级降额 / To derating 1 *)
                eRsn := eIRsnOverTemp;
            END_IF
        eStDer1:                        (* 一级降额相：带回差迁移 / Level 1 with hysteresis *)
            IF (fTempC > fTStopC) OR (fVoltV > fVoltMaxV) THEN
                _eState := eStDer2;
                IF fVoltV > fVoltMaxV THEN
                    eRsn := eIRsnOverVolt;  (* 过压归因 / Over-volt attribution *)
                ELSE
                    eRsn := eIRsnOverTemp;
                END_IF
            ELSIF fTempC < (fT1C - fHysC) THEN
                _eState := eStNormal;   (* 回差解除 / Release by hysteresis *)
            END_IF
        eStDer2:                        (* 二级降额相 / Level 2 *)
            IF (fTempC < fT1C) AND (fVoltV < fVoltMaxV) THEN
                _eState := eStDer1;     (* 双条件回落才降级 / Demote only when both recover *)
            ELSIF fTempC > fTStopC THEN
                _eState := eStStop;     (* 升停机相 / To stop *)
                eRsn := eIRsnOverTemp;  (* 停机相为过温专用 / Stop phase is over-temp only *)
            END_IF
        eStStop:                        (* 停机相：降温回差后回一级 / Stop: recover to level 1 *)
            IF (fTempC < fTStopC - fHysC) AND (fVoltV < fVoltMaxV) THEN
                _eState := eStDer1;
            END_IF
    ELSE
        _eState := eStNormal;           (* ELSE 兜底回 Normal 降级路径 / ELSE fallback to Normal *)
        uCode := 16#0104;               (* 状态越界报码 / Code on illegal state *)
    END_CASE
END_IF

(* === 段 3 · 输出映射与故障码（CASE 内未触碰输出枚举）=== *)
eMode := eMNormal;                      (* 相映射默认 / Default mapping *)
IF _eState = eStDer1 THEN
    eMode := eMDerat1;                  (* 一级降额映射 / Map level 1 *)
ELSIF _eState = eStDer2 THEN
    eMode := eMDerat2;                  (* 二级降额映射 / Map level 2 *)
ELSIF _eState = eStStop THEN
    eMode := eMStop;                    (* 停机映射 / Map stop *)
END_IF
eReason := eRsnNone;                    (* 原因映射默认 / Default reason *)
IF eRsn = eIRsnOverTemp THEN
    eReason := eRsnOverTemp;            (* 过温原因映射 / Map over-temp *)
ELSIF eRsn = eIRsnOverVolt THEN
    eReason := eRsnOverVolt;            (* 过压原因映射 / Map over-volt *)
END_IF
IF (NOT bRun) OR (_eState = eStStop) THEN
    fPowerLimKw := 0.0;                 (* 停机或撤使能封零 / Zero power limit *)
ELSIF _eState = eStDer2 THEN
    fPowerLimKw := fPowerNomKw * DL_IDC_PCT2;   (* 二级限值 [kW] / Level 2 limit *)
ELSIF _eState = eStDer1 THEN
    fPowerLimKw := fPowerNomKw * DL_IDC_PCT1;   (* 一级限值 [kW] / Level 1 limit *)
ELSE
    fPowerLimKw := fPowerNomKw;         (* 额定限值 [kW] / Nominal limit *)
END_IF
bDerating := (_eState = eStDer1) OR (_eState = eStDer2);    (* 降额激活标志 / Derating active *)
bError := (uCode <> 16#0000);           (* 故障标志配对 / Fault flag paired *)
uErrorId := WORD_TO_UDINT(uCode);       (* 码位单点写入（16#0000_0104 形态）/ Single write point *)
END_FUNCTION_BLOCK

(* ---- FB_DL_InverterGridSync.st ---- *)
//==============================================================================
// 功能块：FB_DL_InverterGridSync ｜ 中文名称：逆变器并网同步条件监视
// 所属子库：DL_Device ｜ 版本：v1.0.0 ｜ 兼容：CODESYS V3.5+ / TwinCAT 3 / 汇川 InoProShop
// 功能描述：并网前/并网中同步条件四窗监视：电压幅值窗（网侧三相幅值
//           相对其均值的最大偏差，百分比口径，见边界行为①的窗语义披
//           露）、频率差窗（Hz）、相角差窗（归一 ±180 度）、相序窗
//           （由上游判定给出布尔），四窗全过并持续 tConfirm 才置同步
//           与合闸许可建议。阻塞掩码逐位可观测（电压/频率/相角/相序/
//           输入非法）。仅监视不控合闸（合闸执行由上位断路器逻辑裁
//           决，本件零执行输出）。规格引脚表未提供逆变器侧电压幅值输
//           入，电压窗按「网侧三相幅值相对均值的最大偏差」实现（窗判
//           据不变：偏差超容差即阻塞 bit0），网-逆幅值差需上游增补引
//           脚后切换口径（主动偏离披露，见修订历史）。
// 开源溯源 (Origin)：道莅原创实现（参考 并网同步条件公开工程惯例（电压/频率/相角/相序四窗） 分类与参数域）
// 单位表：电压[V] / 频率[Hz] / 相角[度] / 电压偏差[%] / 容差[%/Hz/度] / 确认延时[ms]
// 错误码表：16#0003_0190 信息级（网侧或逆变侧频率小于等于 0：断线/停机，
//           频率差不判，不置 bError）/ 16#0003_0191 信息级（相角差跨
//           ±180 度发生归一，提示原始差超出半圆，不置 bError）/
//           16#0003_0369 故障级（任一输入非有限，置 bError）/
//           16#0003_036A 故障级（容差组态非法：电压/频率容差非正或相
//           角容差非正、不小于 180 度，置 bError）/ 16#0003_036B 故障
//           级兜底（状态机落 ELSE 或非法状态，置 bError 并撤许可）
// 状态机：E_DL_GridSyncState（eIdle=0 / eChecking=10 / eConfirmed=20 /
//           eFault=99），CASE 含 ELSE 兜底，ELSE 置 036B 并撤许可、
//           全掩码置位（安全侧 = 合闸许可绝不残留）
// 边界行为：① 电压窗语义披露：fVoltDiffPct = max|V相 − V均值| / |V均值|
//           乘 100（三相幅值偏差窗）；V 均值绝对值小于容差（断线/无
//           压）→ 偏差置 0 且窗判失败阻塞 bit0，不做除法；② 相角差
//           归一用条件加减循环（禁 MOD：负数取余三平台不一致，R10 家
//           族），WHILE 带防死锁计数器（上限 4 次迭代），归一后仍出
//           ±180 度 → 相角窗判失败阻塞 bit2；归一发生 → 信息 0191；
//           ③ 任一输入非有限（NaN 自反判 + Inf 幅值上限判，R79）→ 故
//           障 0369 + 掩码 bit4 + bPermitClose := FALSE；④ 网侧或逆变
//           侧频率小于等于 0 → 信息 0190，频率差不判（防除零/防伪同
//           步），掩码 bit1；⑤ 相序不 OK → 掩码 bit3；⑥ 容差组态非
//           法 → 故障 036A + 掩码 bit4；⑦ 失能 → bPermitClose :=
//           FALSE（R72）、bSyncOk := FALSE、回 eIdle；⑧ 确认定时器
//           无条件周期刷新，四窗任一失守即时撤许可并回 eChecking
//           （许可是逐拍实时判定，不锁存）。
// 修订历史：v1.0.0 2026-11-17 首版（R25 派单 · §4.4）
//==============================================================================
(*------------------------------------------------------------------------------
 * 枚举: E_DL_GridSyncState（归属 DL_Device，与 FB_DL_InverterGridSync 同文件）
 *----------------------------------------------------------------------------*)
TYPE E_DL_GridSyncState :
(
    eIdle      := 0,   // 失能/待机：许可撤、掩码全零待刷新 / Idle: permit withdrawn, mask pending refresh
    eChecking  := 10,  // 四窗评估中：确认延时未满 / Checking: windows evaluated, confirm timer running
    eConfirmed := 20,  // 同步确认：四窗全过且持续满 tConfirm / Confirmed: all windows passed for tConfirm
    eFault     := 99   // 故障兜底态：非有限/组态非法/非法状态 / Fault fallback
);
END_TYPE
FUNCTION_BLOCK FB_DL_InverterGridSync
VAR_INPUT
    afGridVoltV  : ARRAY[0..2] OF LREAL;       // 网侧三相电压幅值 [V] / Grid three-phase voltage magnitudes [V]
    fGridFreqHz  : LREAL;                      // 网侧频率 [Hz] / Grid frequency [Hz]
    fInvFreqHz   : LREAL;                      // 逆变侧频率 [Hz] / Inverter frequency [Hz]
    fGridPhaseDeg : LREAL;                     // 网侧相角 [度] / Grid phase angle [deg]
    fInvPhaseDeg : LREAL;                      // 逆变侧相角 [度] / Inverter phase angle [deg]
    fVoltTolPct  : LREAL := 10.0;              // 电压窗容差 [百分数] / Voltage window tolerance [percent]
    fFreqTolHz   : LREAL := 0.2;               // 频率窗容差 [Hz] / Frequency window tolerance [Hz]
    fPhaseTolDeg : LREAL := 10.0;              // 相角窗容差 [度]，域 0~180 开区间 / Phase window tolerance [deg], domain 0..180 open
    tConfirm     : TIME := T#2S;               // 同步确认延时 [ms] / Sync confirmation delay [ms]
    bPhaseSeqOk  : BOOL;                       // 相序判定结果，由上游给出 / Phase-sequence verdict, given by upstream
    bEnable      : BOOL;                       // 总使能 / Master enable
    bReset       : BOOL;                       // 复位，上升沿清状态与掩码 / Reset, rising edge clears state and mask
END_VAR
VAR_OUTPUT
    bSyncOk      : BOOL;                       // 四窗全过且确认延时满 / All windows passed and confirmed
    bPermitClose : BOOL;                       // 合闸许可建议，只读语义，仅监视不控合闸 / Close-permit suggestion, read-only semantics
    fVoltDiffPct : LREAL;                      // 电压幅值偏差 [百分数]（三相幅值偏差窗口径）/ Voltage deviation [percent], three-phase deviation window
    fFreqDiffHz  : LREAL;                      // 频率差 [Hz]，频率无效时保持 0 / Frequency difference [Hz], zero when invalid
    fPhaseDiffDeg : LREAL;                     // 相角差 [度]，已归一 ±180 / Phase difference [deg], normalized to plus-minus 180
    uBlockMask   : WORD;                       // 阻塞掩码：bit0 电压 / bit1 频率 / bit2 相角 / bit3 相序 / bit4 输入或组态非法 / Block mask bits
    eErr         : UDINT;                      // 错误码，0 = 无错，码位 16#0003_0190 起信息级、16#0003_0369 起故障级（分带见错误码表） / Error code, 0 = no error, band info/fault per the code table
    bError       : BOOL;                       // 故障级标志，仅故障级错误置位 / Fault-class flag, set only on fault-level codes
    bValid       : BOOL;                       // 监视数据可用标志，失能/故障闸显式 FALSE / Monitoring usable flag, explicit FALSE on disable/fault gates
    eState       : E_DL_GridSyncState;         // 主状态机当前状态 / Current state of the main state machine
END_VAR
VAR
    fbReset      : R_TRIG;                     // 复位上升沿检测实例 / Reset rising edge detector
    fbConfirm    : TON;                        // 同步确认定时器 / Sync confirmation timer
    fVoltAvg     : LREAL;                      // 三相电压均值 [V] / Mean of three-phase voltages [V]
    fVoltDev     : LREAL;                      // 当前相电压偏差绝对值 [V] / Absolute deviation of current phase [V]
    fVoltDevMax  : LREAL;                      // 三相最大偏差绝对值 [V] / Max absolute deviation across phases [V]
    uPh          : INT;                        // 相循环索引 [—] / Phase loop index
    fPhaseRaw    : LREAL;                      // 归一前相角差 [度] / Raw phase difference before normalization [deg]
    nNormGuard   : INT;                        // 归一循环防死锁计数器 [次] / Normalization loop anti-deadlock counter
    bPhaseNorm   : BOOL;                       // 本拍发生 ±180 度归一 / Normalization occurred this scan
    bVoltOk      : BOOL;                       // 电压窗通过 / Voltage window passed
    bFreqOk      : BOOL;                       // 频率窗通过（频率无效时恒假）/ Frequency window passed (always FALSE when invalid)
    bPhaseAngleOk : BOOL;                      // 相角窗独立判据（不含相序）/ Phase-angle window verdict, sequence excluded
    bPhaseOk     : BOOL;                       // 四窗综合判据：相角 ∧ 相序 / Combined window verdict: angle AND sequence
    bFreqValid   : BOOL;                       // 两侧频率均大于 0，频率差可判 / Both frequencies positive, difference judgeable
END_VAR
VAR CONSTANT
    DL_GSY_CODE_INFO_1 : UDINT := 16#0003_0190;   // 信息级槽 1（频率小于等于 0） / info slot 1
    DL_GSY_CODE_INFO_2 : UDINT := 16#0003_0191;   // 信息级槽 2（相角差归一提示） / info slot 2
    DL_GSY_CODE_FLT_1  : UDINT := 16#0003_0369;   // 故障级槽 1（输入非有限） / fault slot 1
    DL_GSY_CODE_FLT_2  : UDINT := 16#0003_036A;   // 故障级槽 2（容差组态非法） / fault slot 2
    DL_GSY_CODE_FLT_3  : UDINT := 16#0003_036B;   // 故障级槽 3（非法状态兜底） / fault slot 3, illegal-state fallback
    DL_GS_ZERO   : LREAL := 0.0;               // 零值常量，避免裸字面量 [—] / Zero constant, avoids a bare literal
    DL_GS_EPS    : LREAL := 1.0E-6;            // 浮点比较容差 [—] / Float comparison tolerance
    DL_GS_INF    : LREAL := 1.7976931348623157E308;  // LREAL 幅值上限，Inf 判据 / LREAL magnitude ceiling, Inf criterion
    DL_GS_HALF   : LREAL := 180.0;             // 相角归一半圆 [度] / Phase normalization half-circle [deg]
    DL_GS_FULL   : LREAL := 360.0;             // 相角整圆 [度] / Phase full circle [deg]
    DL_GS_NORM_MAX : INT := 4;                 // 归一循环最大迭代 [次]，防死锁 / Normalization loop max iterations, anti-deadlock
    DL_GS_BIT0   : WORD := 16#0001;            // 掩码 bit0：电压窗 / mask bit 0: voltage window
    DL_GS_BIT1   : WORD := 16#0002;            // 掩码 bit1：频率窗 / mask bit 1: frequency window
    DL_GS_BIT2   : WORD := 16#0004;            // 掩码 bit2：相角窗 / mask bit 2: phase window
    DL_GS_BIT3   : WORD := 16#0008;            // 掩码 bit3：相序窗 / mask bit 3: phase-sequence window
    DL_GS_BIT4   : WORD := 16#0010;            // 掩码 bit4：输入或组态非法 / mask bit 4: input or config illegal
END_VAR

(*------------------------------------------------------------------------------
 * 段 1｜无条件刷新区（红线 5）：复位沿检测在任何分支之外周期调用
 *----------------------------------------------------------------------------*)
fbReset(CLK := bReset);                        // 复位沿检测无条件刷新 / reset edge refreshed unconditionally

(*------------------------------------------------------------------------------
 * 段 2｜复位沿处理（改写置于沿后，防吞沿 R39）
 *----------------------------------------------------------------------------*)
IF fbReset.Q THEN
    eState       := E_DL_GridSyncState.eIdle;
    eErr         := 16#0000_0000;              // 复位清码 / reset clears code
    bError       := FALSE;                     // 复位清故障 / reset clears fault
    uBlockMask   := 16#0000;                   // 掩码清零 / mask zeroed
    bSyncOk      := FALSE;                     // 同步撤 / sync withdrawn
    bPermitClose := FALSE;                     // 许可撤（安全侧）/ permit withdrawn, safe side
    bValid       := FALSE;                     // 可用撤 / usable withdrawn
END_IF

(*------------------------------------------------------------------------------
 * 段 3｜非有限输入闸（三相电压 + 四标量：NaN 自反判 + Inf 幅值上限判，R79）
 *----------------------------------------------------------------------------*)
IF (afGridVoltV[0] <> afGridVoltV[0]) OR (ABS(afGridVoltV[0]) >= DL_GS_INF)
   OR (afGridVoltV[1] <> afGridVoltV[1]) OR (ABS(afGridVoltV[1]) >= DL_GS_INF)
   OR (afGridVoltV[2] <> afGridVoltV[2]) OR (ABS(afGridVoltV[2]) >= DL_GS_INF)
   OR (fGridFreqHz <> fGridFreqHz) OR (ABS(fGridFreqHz) >= DL_GS_INF)
   OR (fInvFreqHz <> fInvFreqHz) OR (ABS(fInvFreqHz) >= DL_GS_INF)
   OR (fGridPhaseDeg <> fGridPhaseDeg) OR (ABS(fGridPhaseDeg) >= DL_GS_INF)
   OR (fInvPhaseDeg <> fInvPhaseDeg) OR (ABS(fInvPhaseDeg) >= DL_GS_INF) THEN
    eState       := E_DL_GridSyncState.eFault;
    eErr         := DL_GSY_CODE_FLT_1;         // 故障级：任一输入非有限 / fault: non-finite input
    bError       := TRUE;                      // 故障级必置 bError（R45 配对）/ fault-class pairs with bError
    bValid       := FALSE;                     // 输出不可用 / outputs unusable
    bSyncOk      := FALSE;                     // 同步撤 / sync withdrawn
    bPermitClose := FALSE;                     // 许可撤（R72，安全侧）/ permit withdrawn, safe side
    uBlockMask   := DL_GS_BIT4;                // 掩码 bit4：输入非法 / mask bit 4: input illegal
    fVoltDiffPct := DL_GS_ZERO;                // 偏差出口清零 / deviation outputs zeroed
    fFreqDiffHz  := DL_GS_ZERO;                // 偏差出口清零 / deviation outputs zeroed
    fPhaseDiffDeg := DL_GS_ZERO;               // 偏差出口清零 / deviation outputs zeroed
    fbConfirm(IN := FALSE, PT := tConfirm);    // 确认定时器断输入（无条件调用保持）/ confirm timer input broken, still called
    RETURN;
END_IF

(*------------------------------------------------------------------------------
 * 段 4｜容差组态闸（电压/频率容差非正、相角容差非正或不小于 180 度）
 *----------------------------------------------------------------------------*)
IF (fVoltTolPct <= DL_GS_EPS) OR (fFreqTolHz <= DL_GS_EPS)
   OR (fPhaseTolDeg <= DL_GS_EPS) OR (fPhaseTolDeg >= DL_GS_HALF) THEN
    eState       := E_DL_GridSyncState.eFault;
    eErr         := DL_GSY_CODE_FLT_2;         // 故障级：容差组态非法 / fault: tolerance config invalid
    bError       := TRUE;                      // 故障级必置 bError（R45 配对）/ fault-class pairs with bError
    bValid       := FALSE;                     // 输出不可用 / outputs unusable
    bSyncOk      := FALSE;                     // 同步撤 / sync withdrawn
    bPermitClose := FALSE;                     // 许可撤（R72，安全侧）/ permit withdrawn, safe side
    uBlockMask   := DL_GS_BIT4;                // 掩码 bit4：组态非法 / mask bit 4: config illegal
    fbConfirm(IN := FALSE, PT := tConfirm);    // 确认定时器断输入（无条件调用保持）/ confirm timer input broken, still called
    RETURN;
END_IF

(*------------------------------------------------------------------------------
 * 段 5｜四窗评估（电压/频率/相角/相序），先算窗口再刷定时器（定时器无条件调用）
 *----------------------------------------------------------------------------*)
(*--- 5.1 电压窗：三相幅值相对均值最大偏差（见边界行为①口径披露）---*)
fVoltAvg := (afGridVoltV[0] + afGridVoltV[1] + afGridVoltV[2]) / 3.0;  // 三相均值 [V] / three-phase mean [V]
fVoltDevMax := DL_GS_ZERO;                     // 最大偏差复位 / max deviation reset
FOR uPh := 0 TO 2 DO
    fVoltDev := ABS(afGridVoltV[uPh] - fVoltAvg);  // 当前相偏差绝对值 [V] / current phase deviation [V]
    IF fVoltDev > fVoltDevMax THEN
        fVoltDevMax := fVoltDev;               // 保留最大 / keep the max
    END_IF
END_FOR
IF ABS(fVoltAvg) > DL_GS_EPS THEN
    fVoltDiffPct := fVoltDevMax / ABS(fVoltAvg) * 100.0;  // 相对偏差百分比口径，除子已判 / relative deviation, divisor checked
    bVoltOk := fVoltDiffPct <= fVoltTolPct;    // 窗判 / window verdict
ELSE
    fVoltDiffPct := DL_GS_ZERO;                // 无压/断线：偏差不可算，置 0 / no voltage: deviation not computable, zeroed
    bVoltOk := FALSE;                          // 窗判失败 / window fails
END_IF

(*--- 5.2 频率窗：两侧频率大于 0 才判差（信息 0190，防伪同步）---*)
IF (fGridFreqHz > DL_GS_EPS) AND (fInvFreqHz > DL_GS_EPS) THEN
    bFreqValid := TRUE;                        // 频率差可判 / difference judgeable
    fFreqDiffHz := fInvFreqHz - fGridFreqHz;   // 频率差 [Hz] / frequency difference [Hz]
    bFreqOk := ABS(fFreqDiffHz) <= fFreqTolHz; // 窗判 / window verdict
ELSE
    bFreqValid := FALSE;                       // 频率无效：断线/停机 / frequency invalid: offline or stopped
    fFreqDiffHz := DL_GS_ZERO;                 // 频率差出口清零 / difference output zeroed
    bFreqOk := FALSE;                          // 频率差不判，窗判失败 / difference not judged, window fails
END_IF

(*--- 5.3 相角窗：条件加减归一 ±180 度（禁 MOD，R10 家族；WHILE 防死锁计数器）---*)
fPhaseRaw := fInvPhaseDeg - fGridPhaseDeg;     // 归一前相角差 [度] / raw phase difference [deg]
fPhaseDiffDeg := fPhaseRaw;                    // 归一工作副本 / working copy
nNormGuard := 0;                               // 防死锁计数清零 / anti-deadlock counter zeroed
WHILE ((fPhaseDiffDeg > DL_GS_HALF) OR (fPhaseDiffDeg < -DL_GS_HALF)) AND (nNormGuard < DL_GS_NORM_MAX) DO
    IF fPhaseDiffDeg > DL_GS_HALF THEN
        fPhaseDiffDeg := fPhaseDiffDeg - DL_GS_FULL;   // 越上半圆减整圆 / above half-circle subtract full circle
    ELSE
        fPhaseDiffDeg := fPhaseDiffDeg + DL_GS_FULL;   // 越下半圆加整圆 / below half-circle add full circle
    END_IF
    nNormGuard := nNormGuard + 1;              // 迭代计数 / iteration count
END_WHILE
bPhaseNorm := ABS(fPhaseRaw) > DL_GS_HALF;     // 原始差超半圆即发生归一 / normalization occurred when raw beyond half-circle
bPhaseAngleOk := (ABS(fPhaseDiffDeg) <= fPhaseTolDeg) AND (nNormGuard < DL_GS_NORM_MAX);  // 相角窗独立判，归一失败亦判失败 / phase-angle window verdict, failed normalization also fails
bPhaseOk := bPhaseAngleOk AND bPhaseSeqOk;     // 四窗综合判：相角 ∧ 相序 / combined window verdict: angle AND sequence

(*--- 5.5 确认定时器：无条件周期刷新（红线 5）---*)
fbConfirm(IN := bEnable AND bVoltOk AND bFreqOk AND bPhaseOk,  // 四窗全过且使能才计时 / timer runs when enabled and all windows pass
          PT := tConfirm);                     // 确认延时 / confirmation delay

(*------------------------------------------------------------------------------
 * 段 6｜阻塞掩码逐拍装配（先清后置，逐位可观测）
 *----------------------------------------------------------------------------*)
uBlockMask := 16#0000;                         // 掩码逐拍重装配 / mask reassembled per scan
IF NOT bVoltOk THEN
    uBlockMask := uBlockMask OR DL_GS_BIT0;    // bit0：电压窗 / bit 0: voltage window
END_IF
IF NOT bFreqOk THEN
    uBlockMask := uBlockMask OR DL_GS_BIT1;    // bit1：频率窗（含频率无效）/ bit 1: frequency window, incl. invalid
END_IF
IF NOT bPhaseAngleOk THEN
    uBlockMask := uBlockMask OR DL_GS_BIT2;    // bit2：相角窗（含归一失败）/ bit 2: phase-angle window
END_IF
IF NOT bPhaseSeqOk THEN
    uBlockMask := uBlockMask OR DL_GS_BIT3;    // bit3：相序窗 / bit 3: phase-sequence window
END_IF

(*------------------------------------------------------------------------------
 * 段 7｜状态机：CASE 含 ELSE 兜底（非法状态 → 036B + 撤许可，安全侧）
 *----------------------------------------------------------------------------*)
CASE eState OF

    E_DL_GridSyncState.eIdle:
        bValid := FALSE;                       // 失能闸显式不可用（R72）/ explicit FALSE on disable gate
        bSyncOk := FALSE;                      // 同步撤 / sync withdrawn
        bPermitClose := FALSE;                 // 许可撤（安全侧）/ permit withdrawn, safe side
        eErr := 16#0000_0000;                  // 待机无错 / no error in idle
        bError := FALSE;                       // 待机无故障 / no fault in idle
        IF bEnable THEN
            eState := E_DL_GridSyncState.eChecking;    // 使能进评估 / enable enters checking
        END_IF

    E_DL_GridSyncState.eChecking:
        IF NOT bEnable THEN
            eState := E_DL_GridSyncState.eIdle;        // 失能回待机 / disable returns to idle
            bValid := FALSE;                   // 失能闸显式不可用 / explicit FALSE on disable gate
            bPermitClose := FALSE;             // 许可撤（安全侧）/ permit withdrawn, safe side
            bSyncOk := FALSE;                  // 同步撤 / sync withdrawn
        ELSE
            bValid := TRUE;                    // 评估态监视数据可用 / monitoring usable in checking
            eErr := 16#0000_0000;              // 评估态先清码 / checking clears code first
            IF bPhaseNorm THEN
                eErr := DL_GSY_CODE_INFO_2;    // 信息级：相角差跨 ±180 度归一 / info: phase normalized across half-circle
            END_IF
            IF NOT bFreqValid THEN
                eErr := DL_GSY_CODE_INFO_1;    // 信息级：频率无效优先于归一提示 / info: invalid frequency outranks normalization hint
            END_IF
            bError := FALSE;                   // 信息级不置 bError / info never raises bError
            bSyncOk := FALSE;                  // 未确认前同步撤 / sync withdrawn before confirmation
            bPermitClose := FALSE;             // 未确认前许可撤 / permit withdrawn before confirmation
            IF fbConfirm.Q THEN
                eState := E_DL_GridSyncState.eConfirmed;   // 确认延时满进确认态 / delay elapsed enters confirmed
            END_IF
        END_IF

    E_DL_GridSyncState.eConfirmed:
        IF NOT bEnable THEN
            eState := E_DL_GridSyncState.eIdle;
            bValid := FALSE;
            bPermitClose := FALSE;             // 许可撤（安全侧）/ permit withdrawn, safe side
            bSyncOk := FALSE;
        ELSE
            bValid := TRUE;                    // 确认态监视数据可用 / monitoring usable in confirmed
            eErr := 16#0000_0000;              // 先清码 / clear code first
            IF bPhaseNorm THEN
                eErr := DL_GSY_CODE_INFO_2;    // 信息级：归一提示 / info: normalization hint
            END_IF
            IF NOT bFreqValid THEN
                eErr := DL_GSY_CODE_INFO_1;    // 信息级：频率无效优先 / info: invalid frequency outranks
            END_IF
            bError := FALSE;                   // 信息级不置 bError / info never raises bError
            bSyncOk := fbConfirm.Q;            // 同步逐拍实时判定，不锁存 / sync judged per scan, not latched
            bPermitClose := fbConfirm.Q AND bFreqValid;  // 许可逐拍实时判定，频率无效不许可 / permit judged per scan, invalid frequency blocks
            IF NOT fbConfirm.Q THEN
                eState := E_DL_GridSyncState.eChecking;    // 四窗任一失守回评估（定时器自动重启）/ any window lost returns to checking
            END_IF
        END_IF

    ELSE
        eState := E_DL_GridSyncState.eFault;   // 非法状态兜底 / illegal-state fallback
        eErr   := DL_GSY_CODE_FLT_3;           // 故障级兜底：非法状态 / fault fallback: illegal state
        bError := TRUE;                        // 故障级必置 bError / fault-class pairs with bError
        bValid := FALSE;                       // 输出不可用 / outputs unusable
        bSyncOk := FALSE;                      // 同步撤 / sync withdrawn
        bPermitClose := FALSE;                 // 许可撤（安全侧，绝不残留）/ permit withdrawn, never residual
END_CASE
END_FUNCTION_BLOCK

(* ---- FB_DL_InverterPdiPoll.st ---- *)
(*
  FB_DL_InverterPdiPoll  —  逆变器 PDI 参数周期读取（单拍单发 + 站表台账） / Inverter PDI parameter cyclic poll with a station ledger
  分类 Category : DL_Device
  版本 Version  : 1.0.0
  来源 Source   : t1-7-plcnext — PDI 应用族零检索深化（基于 PdiReadScheduler 底座）
  溯源 Origin   : clean-room 实现，未复制任何源码行
  功能 Function : 1) 站表 aSlot 逐站轮询：eIdle（间隔到）→ eReq（单发 bStart）→ eWait
                  （等 bDone）→ eJudge（读-比-判：bSuccess 且 uActLen = 期望长度）；
                  2) 单拍单发纪律：全轮询任意时刻仅一个在途请求（状态机单相承载）；
                  3) 台账：uOkTotal / uFailTotal / 站内连续失败计数，达 nFailLatch 阈
                  → 故障级 03FD 锁存；
                  4) 站间推进沿 041C；全站巡检一周完成沿 041D；连续失败未达阈提示 041E。
  边界 Boundary : ① 组态闸：uStationCnt < 1 或 > 8 → 03FC 锁存（站表容量下限 >= 1）；
                  ② Device 段 0003 故障带仅余 03FC~03FF，本件启用 03FC/03FD 两格，
                  分段理由：03xx 带收口分配，不足溢出走 05xx 副带（本轮未占用）；
                  ③ fbPdi 输入引脚在 eIdle 相整定、eReq 相单发，禁批量并发；
                  ④ 无 GVL 依赖：纯引脚输入输出，无外部变量引用，无物理 IO 地址。
  依赖 Depends  : FB_DL_PdiReadScheduler（注入，不实例化，引脚按 registry 实名）；Standard.library（TON / R_TRIG）
  码表 Error codes（Device 段 0003，窗口 041C~041E / 故障 03FC~03FD）:
    16#0003_03FC 故障级：组态非法（站数界外），锁存至 bReset
    16#0003_03FD 故障级：站点连续失败达阈锁存（台账口径），锁存至 bReset
    16#0003_041C 信息级：站间推进沿（切换下一站）
    16#0003_041D 信息级：全站巡检一周完成沿
    16#0003_041E 信息级：连续失败未达阈提示（伴随态）
  修订历史 Revision :
    2026-11-19  v1.0.0  R41 首版（批次 4 · 序号 1）
*)

TYPE E_DL_InvPollState :
(
    eIdle  := 0,    // 空闲：等站间间隔 / Idle, waiting the inter-station gap
    eReq   := 10,   // 请求：单发启动 / Request, one-shot start
    eWait  := 20,   // 等待：等传输层完成 / Wait, transport completion
    eJudge := 30,   // 判定：读-比-判三段 / Judge, read-compare-verdict
    eFault := 90    // 故障：连续失败锁定 / Fault, latched
);
END_TYPE

FUNCTION_BLOCK FB_DL_InverterPdiPoll
VAR_INPUT
    aSlot        : ARRAY[1..8] OF UINT;   // 站表（设备号）[号] / Station slot table
    uStationCnt  : UINT := 1;         // 站数 [站]，域 1..8 / Station count
    uIndex       : UINT := 16#2035;   // PDI 对象索引（逆变器参数例）/ Object index
    uSubindex    : USINT := 0;        // 对象子索引 / Object subindex
    nExpLen      : INT := 2;          // 期望数据长度 [字节] / Expected data length
    tPollGap     : TIME := T#100MS;   // 站间间隔 [ms]，域 > 0 / Inter-station gap
    tWaitTo      : TIME := T#2S;      // 在途等待超时 [ms]，域 > 0 / In-flight wait timeout
    nFailLatch   : INT := 3;          // 连续失败锁存阈 [次]，域 >= 1 / Consecutive-fail latch threshold
    bEnable      : BOOL := FALSE;     // 轮询使能 [-] / Poll enable
    bReset       : BOOL := FALSE;     // 复位，上升沿清故障锁存 / Reset edge clears fault latch
END_VAR
VAR_IN_OUT
    fbPdi        : FB_DL_PdiReadScheduler;  // PDI 调度底座（注入，不实例化）/ PDI scheduler base
END_VAR
VAR_OUTPUT
    eState       : E_DL_InvPollState; // 状态出口，段尾单点映射 / State outlet
    uCurSlot     : UINT;              // 当前站号出口 [号] / Current slot outlet
    uIdx         : UINT;              // 当前站序号（1 基）[站] / Current station index
    uOkTotal     : UDINT;             // 累计成功数 [次]，饱和不回绕 / Total success count
    uFailTotal   : UDINT;             // 累计失败数 [次]，饱和不回绕 / Total failure count
    bError       : BOOL;              // 故障锁存标志 / Fault latch flag
    nErrId       : UDINT;             // 事件码，0 = 无事件 / Event code
END_VAR
VAR
    tonGap       : TON;               // 站间间隔定时器（自复位口径），无条件刷新 / Inter-station gap timer
    tonWaitTo    : TON;               // 在途等待定时器（专用超时命名），无条件刷新 / In-flight wait timer
    rtReset      : R_TRIG;            // 复位沿实例，无条件刷新 / Reset edge instance
    _eState      : E_DL_InvPollState := E_DL_InvPollState.eIdle;  // 内部相位（CASE 唯一写入目标）/ Internal phase
    _uIdx        : UINT := 1;         // 内部站序号（1 基）/ Internal station index
    _nFailRun    : INT;               // 站内连续失败计数 [次] / Consecutive-fail streak
    _bFault      : BOOL;              // 故障锁存位（锁存量）/ Latched fault bit
    _uFault      : UDINT;             // 故障码锁存（锁存量）/ Latched fault code
    _uInfo       : UDINT;             // 信息码，每拍重算 / Transient info code
END_VAR
VAR CONSTANT
    DL_IPP_CNT_MAX : UDINT := 16#FFFF_FFFE;  // 台账计数饱和上限 [次] / Ledger saturation bound
END_VAR

(* —— 段 0：定时器与沿实例无条件周期刷新（禁置于 IF/CASE 内） —— *)
rtReset(CLK := bReset);                                   // 复位沿（每拍必调）
tonGap(IN := (_eState = E_DL_InvPollState.eIdle) AND bEnable AND (NOT _bFault), PT := tPollGap);
                                                          // 站间间隔（每拍必调，TON 自复位口径 IN 断即清）
tonWaitTo(IN := (_eState = E_DL_InvPollState.eWait), PT := tWaitTo);   // 在途等待（单相独占）

(* —— 段 1：单拍量预清零（锁存量 _bFault/_uFault/台账计数不入清单，禁同拍抹除） —— *)
_uInfo := 16#0000_0000;             // 信息码每拍重算
nErrId := 16#0000_0000;             // 事件码缺省无事件

(* —— 段 2：复位沿 + 组态域闸（当拍量判据） —— *)
IF rtReset.Q THEN                   // rtReset.Q = 当拍量
    _bFault := FALSE;               // 清故障锁存位
    _uFault := 16#0000_0000;        // 清故障锁存码
END_IF
IF (UINT_TO_INT(uStationCnt) < 1) OR (UINT_TO_INT(uStationCnt) > 8)
   OR (TIME_TO_DINT(tPollGap) <= 0) OR (TIME_TO_DINT(tWaitTo) <= 0) OR (nFailLatch < 1) THEN
    _uFault := 16#0003_03FC;        // 故障级：组态非法
    _bFault := TRUE;
END_IF

(* —— 段 3：底座输入整定（每拍写入；bStart 仅 eReq 相电平置位构成单发沿） —— *)
fbPdi.bEnable := bEnable AND (NOT _bFault);   // 底座使能随本件
IF (UINT_TO_INT(_uIdx) >= 1) AND (UINT_TO_INT(_uIdx) <= 8) THEN
    fbPdi.uSlot := aSlot[UINT_TO_INT(_uIdx)]; // 当前站号下装（界内守卫）
END_IF
fbPdi.uIndex := uIndex;             // 对象索引下装
fbPdi.uSubindex := uSubindex;       // 子索引下装
fbPdi.nExpLen := nExpLen;           // 期望长度下装（比较段判据）
fbPdi.bStart := (_eState = E_DL_InvPollState.eReq);   // 单发沿（eReq 单相电平，下一相即断）

(* —— 段 4：相位机（CASE 全覆盖 + ELSE 兜底；单拍单发由状态机单相承载） —— *)
CASE _eState OF

E_DL_InvPollState.eIdle:
    IF _bFault THEN
        _eState := E_DL_InvPollState.eFault;    // 故障相
    ELSIF bEnable AND tonGap.Q THEN
        fbPdi.bEnable := TRUE;                  // 底座使能确认
        _eState := E_DL_InvPollState.eReq;      // 进请求相（bStart 下一拍电平置位成沿）
    END_IF

E_DL_InvPollState.eReq:
    IF _bFault THEN
        _eState := E_DL_InvPollState.eFault;    // 故障相（bStart 已断）
    ELSE
        _eState := E_DL_InvPollState.eWait;     // bStart 单发即进等待相（下一拍电平断）
    END_IF

E_DL_InvPollState.eWait:
    IF _bFault THEN
        _eState := E_DL_InvPollState.eFault;    // 故障相
    ELSIF tonWaitTo.Q THEN
        _nFailRun := _nFailRun + 1;             // 超时按失败入账
        uFailTotal := uFailTotal + 1;           // 台账累加
        IF uFailTotal >= DL_IPP_CNT_MAX THEN
            uFailTotal := DL_IPP_CNT_MAX;       // 台账饱和防回绕
        END_IF
        _eState := E_DL_InvPollState.eIdle;     // 回空闲（下一站间隔后重试）
    ELSIF fbPdi.bDone THEN
        _eState := E_DL_InvPollState.eJudge;    // 完成沿：进判定相
    END_IF

E_DL_InvPollState.eJudge:
    IF _bFault THEN
        _eState := E_DL_InvPollState.eFault;    // 故障相
    ELSIF fbPdi.bSuccess AND (fbPdi.uActLen = INT_TO_UINT(nExpLen)) THEN
        uOkTotal := uOkTotal + 1;               // 台账成功累加
        IF uOkTotal >= DL_IPP_CNT_MAX THEN
            uOkTotal := DL_IPP_CNT_MAX;         // 台账饱和防回绕
        END_IF
        _nFailRun := 0;                         // 连败计数清零
        _uInfo := 16#0003_041C;                 // 信息级：站间推进沿（成功随行）
        _uIdx := _uIdx + 1;                     // 下一站
        IF UINT_TO_INT(_uIdx) > UINT_TO_INT(uStationCnt) THEN
            _uIdx := 1;                         // 站表回卷
            _uInfo := 16#0003_041D;             // 信息级：全站巡检一周完成
        END_IF
        _eState := E_DL_InvPollState.eIdle;     // 回空闲
    ELSE
        _nFailRun := _nFailRun + 1;             // 失败或长度不匹配：连败入账
        uFailTotal := uFailTotal + 1;           // 台账累加
        IF uFailTotal >= DL_IPP_CNT_MAX THEN
            uFailTotal := DL_IPP_CNT_MAX;       // 台账饱和防回绕
        END_IF
        IF _nFailRun >= nFailLatch THEN
            _uFault := 16#0003_03FD;            // 故障级：连续失败达阈锁存
            _bFault := TRUE;
            _eState := E_DL_InvPollState.eFault;
        ELSE
            _uInfo := 16#0003_041E;             // 信息级：连败未达阈提示
            _eState := E_DL_InvPollState.eIdle; // 回空闲重试
        END_IF
    END_IF

E_DL_InvPollState.eFault:
    ;                                   // 故障相：等复位沿（段 2 承载迁出）

ELSE
    _uFault := 16#0003_03FC;            // 故障级：非法相位兜底（归并组态码，头注释②）
    _bFault := TRUE;
    _eState := E_DL_InvPollState.eFault;    // 强制回故障相

END_CASE

(* —— 段 5：出口单点映射（名实同源；锁存码回放，禁同拍抹除） —— *)
uCurSlot := aSlot[UINT_TO_INT(_uIdx)];      // 当前站号出口（站表 1..8 静态界内）
IF UINT_TO_INT(_uIdx) < 1 THEN
    uIdx := 1;                      // 序号下界防御
ELSIF UINT_TO_INT(_uIdx) > 8 THEN
    uIdx := 8;                      // 序号上界防御
ELSE
    uIdx := _uIdx;                  // 序号直通
END_IF
IF _bFault THEN
    nErrId := _uFault;              // 故障锁存码回放
ELSE
    nErrId := _uInfo;               // 信息码
END_IF
bError := _bFault;                  // 故障标志与锁存位同源
eState := _eState;                  // 状态出口单点映射

END_FUNCTION_BLOCK

(* ---- FB_DL_IoLinkPortDiag.st ---- *)
(*
  道莅工业代码库 | DL_Device | FB_DL_IoLinkPortDiag
  版本: 1.0.0 | 日期: 2026-11-23 | 轮次: R75
  开源溯源: self-cleanroom（无外部来源；IO-Link 端口诊断语义，零代码行复制）
  功能: IO-Link 端口诊断聚合——8 端口设备质量码/过程数据有效位逐口判坏与计数，
        主站循环翻转看门狗（tWdTimeout 内无翻转判通信丢失，锁存需复位）。
  兼容性: CODESYS 3.5 / TwinCAT 3 / 汇川 InoProShop；仅依赖标准 TON / R_TRIG / F_TRIG，零厂商私有库
  接口: 输入 aPortQuality（8 端口质量码，0=好）/aPdValid（8 端口 PD 有效）/
        bCycleTog（主站循环翻转输入）/tWdTimeout/bEn/bReset；输出 bAllPortsOk/
        bWdOk/uBadCnt/aPortBad/eState/eCause/bError/nErrId。
  码表: 16#0003_038A 故障级：循环看门狗超时（翻转丢失锁存至复位沿）
        16#0003_0410 信息级：存在坏端口（质量码非零或 PD 无效，当拍重算）
        码段说明：0003 段故障子带 03xx / 信息子带 04xx，槽位经全库实扫空闲。
  边界: ① 数组全部固定上界 [1..8]（零 VLA，R75 口径），下标 1..8 由 FOR 常量界
        证明无越界；
        ② 看门狗：rtTog/ftTog 任一沿喂狗，TON IN := NOT 沿，翻转丢失经去抖
        窗锁存；翻转正常时 IN 周期性落 FALSE 自复位（R188 自复位口径）；
        ③ 端口坏为电平判据（不锁存），信息级每拍重算；看门狗丢失为锁存故障；
        ④ TON/R_TRIG/F_TRIG 段 0 无条件周期刷新；⑤ 零全局耦合。
  邻件比对: ProfinetAlarmDiag（PROFINET vs 本件 IO-Link，协议域不同）。
  修订历史: 2026-11-23 v1.0.0 R75 首版（复杂件批 B3 · C12）
*)

TYPE E_DL_IldState :
(
    eOk        := 0,   // 全端口健康且看门狗正常 | All ports healthy, watchdog ok
    ePortFault := 10,  // 存在坏端口 | At least one bad port
    eWdLost    := 20   // 循环看门狗丢失（锁存） | Cycle watchdog lost, latched
);
END_TYPE

TYPE E_DL_IldCause :
(
    eNone        := 0,  // 无故障 | No cause
    eWdNoToggle  := 1,  // 循环翻转丢失 | Cycle toggle lost
    ePortQuality := 2,  // 端口质量码非零 | Port quality code non-zero
    ePdInvalid   := 3   // 端口过程数据无效 | Port PD invalid
);
END_TYPE

FUNCTION_BLOCK FB_DL_IoLinkPortDiag
VAR_INPUT
    bEn          : BOOL := FALSE;    // 诊断使能 [-] | Diagnostics enable
    aPortQuality : ARRAY[1..8] OF BYTE;   // 每端口设备质量码（0=好）[码] | Per-port device quality code, 0 = good
    aPdValid     : ARRAY[1..8] OF BOOL;   // 每端口过程数据有效 [-] | Per-port process data valid
    bCycleTog    : BOOL := FALSE;    // 主站循环翻转输入（每循环取反）[-] | Master cycle toggle input
    tWdTimeout   : TIME := T#100MS;  // 看门狗超时，域 > T#0S | Watchdog timeout
    bReset       : BOOL := FALSE;    // 复位命令，上升沿清锁存 [-] | Reset command, rising edge
END_VAR
VAR_OUTPUT
    bAllPortsOk : BOOL;             // 全端口健康且看门狗正常 [-] | All ports ok and watchdog ok
    bWdOk       : BOOL;             // 循环看门狗正常 [-] | Cycle watchdog ok
    uBadCnt     : UINT;             // 坏端口计数 [口] | Bad port count
    aPortBad    : ARRAY[1..8] OF BOOL;   // 每端口坏标志 [-] | Per-port bad flag
    eState      : E_DL_IldState;    // 状态出口 | State outlet
    eCause      : E_DL_IldCause;    // 成因出口 | Cause outlet
    bError      : BOOL;             // 故障锁存标志 [-] | Fault latch flag
    nErrId      : UDINT;            // 事件码，0 = 无事件 | Event code, 0 = none
END_VAR
VAR
    _bWdLatch : BOOL;               // 看门狗丢失锁存位 | Watchdog lost latch bit
    _eCause   : E_DL_IldCause := E_DL_IldCause.eNone;   // 成因锁存 | Latched cause
    _ePortCau : E_DL_IldCause := E_DL_IldCause.eNone;   // 端口成因当拍归因 | Port cause attribution this scan
    _nBad     : INT;                // 坏端口计数当拍量 [口] | Bad port count this scan
    _bAnyBad  : BOOL;               // 存在坏端口当拍量 [-] | Any bad port this scan
    i         : INT;                // 端口游标（1..8 常量界）| Port cursor, constant bounds
    rtTog     : R_TRIG;             // 翻转上升沿实例，段 0 无条件刷新 | Toggle rising edge instance
    ftTog     : F_TRIG;             // 翻转下降沿实例，段 0 无条件刷新 | Toggle falling edge instance
    rtReset   : R_TRIG;             // 复位沿实例，段 0 无条件刷新 | Reset edge instance
    tonWd     : TON;                // 看门狗计时（喂狗自复位），段 0 无条件刷新 | Watchdog timer, fed by edges
END_VAR

(* —— 段 0：沿与定时器实例无条件周期刷新（R7 红线） —— *)
rtTog(CLK := bCycleTog);                    // 翻转上升沿每拍必调 / Rising edge every scan
ftTog(CLK := bCycleTog);                    // 翻转下降沿每拍必调 / Falling edge every scan
tonWd(IN := NOT (rtTog.Q OR ftTog.Q), PT := tWdTimeout);   // 喂狗：任一沿 IN 落假自复位（边界②）/ Fed by any edge, self-reset
rtReset(CLK := bReset);                     // 复位沿每拍必调 / Reset edge every scan

(* —— 段 1：复位沿 + 看门狗锁存 —— *)
IF rtReset.Q THEN
    _bWdLatch := FALSE;                     // 清看门狗锁存位 / Clear watchdog latch
    _eCause := E_DL_IldCause.eNone;         // 清成因 / Clear cause
END_IF
IF bEn AND tonWd.Q AND (NOT _bWdLatch) THEN
    _bWdLatch := TRUE;                      // 翻转丢失超时锁存 / Toggle loss timeout latch
    _eCause := E_DL_IldCause.eWdNoToggle;   // 归因翻转丢失 / Cause: toggle lost
END_IF

(* —— 段 2：逐端口判坏与计数（下标 1..8 常量界，无越界路径） —— *)
_nBad := 0;                                 // 计数当拍量预清 / Count preset
_bAnyBad := FALSE;                          // 坏标志预清 / Any-bad preset
_ePortCau := E_DL_IldCause.eNone;           // 端口成因预清 / Port cause preset
FOR i := 1 TO 8 DO
    IF (aPortQuality[i] <> 0) OR (NOT aPdValid[i]) THEN
        aPortBad[i] := TRUE;                // 端口坏：质量码非零或 PD 无效 / Port bad by quality or PD
        _nBad := _nBad + 1;                 // 坏端口计数 / Count increment
        _bAnyBad := TRUE;                   // 存在坏端口 / Any bad flag
        IF NOT aPdValid[i] THEN
            _ePortCau := E_DL_IldCause.ePdInvalid;      // 归因 PD 无效（先到先归因）/ Cause: PD invalid
        ELSE
            _ePortCau := E_DL_IldCause.ePortQuality;    // 归因质量码 / Cause: quality code
        END_IF
    ELSE
        aPortBad[i] := FALSE;               // 端口好 / Port good
    END_IF
END_FOR

(* —— 段 3：出口单点映射（名实同源；锁存码回放 + 信息码重算） —— *)
bWdOk := (NOT tonWd.Q) AND (NOT _bWdLatch);              // 看门狗正常判据（锁存后保持坏）/ Watchdog ok judgement
uBadCnt := INT_TO_UINT(_nBad);                           // 坏端口计数出口 / Bad count outlet
bAllPortsOk := (NOT _bWdLatch) AND (_nBad = 0);          // 总健康判据 / All-ok judgement
IF _bWdLatch THEN
    eState := E_DL_IldState.eWdLost;                     // 看门狗丢失态 / Watchdog lost state
ELSIF bEn AND _bAnyBad THEN
    eState := E_DL_IldState.ePortFault;                  // 坏端口态 / Port fault state
ELSE
    eState := E_DL_IldState.eOk;                         // 健康态 / Ok state
END_IF
IF _bWdLatch THEN
    eCause := _eCause;                                   // 锁存成因出口（看门狗）/ Latched watchdog cause
ELSE
    eCause := _ePortCau;                                 // 当拍端口成因出口 / Per-scan port cause
END_IF
bError := _bWdLatch;                                     // 故障标志同源 / Error flag from latch
IF _bWdLatch THEN
    nErrId := 16#0003_038A;                              // 看门狗锁存码回放 / Replay watchdog latch code
ELSIF _bAnyBad THEN
    nErrId := 16#0003_0410;                              // 信息级：存在坏端口（每拍重算）/ Info: bad port present
ELSE
    nErrId := 16#0000_0000;                              // 无事件 / No event
END_IF

END_FUNCTION_BLOCK

(* ---- FB_DL_IonizerAirflowInterlock.st ---- *)
(*
  ==================================================================
  组件名 Component  : FB_DL_IonizerAirflowInterlock
  分类   Category   : DL_Device
  复杂度 Complexity  : cx4
  版本   Version    : 1.0.0
  功能   Purpose    : 离子风机风速联锁。风速低于下限持续 tConfirm 确认窗才锁存
                      （单拍毛刺不动作）；放行门控出口（bPermitOk）与消电离
                      有效性出口（bIonValid）分离；失能即解锁回空闲且输出
                      安全侧断开放行。
  来源   Source     : self-esc（ROADMAP R56 评估项转正；借鉴 ISA-TR84 风量联锁
                      确认窗纪律，clean-room 自研实现，未复制任何文档代码行）
  溯源   Origin     : IEC 61131-3 标准语义的道莅防御性实现；离子风机风速下限
                      联锁为公开防静电工艺语义。
  平台   Platform   : 纯 IEC 61131-3（Standard.library: TON / R_TRIG，无私有库）
  分工声明 Split     : 与 FB_DL_EsdGroundMonitor（接地判级）分工——本件只做
                      风速联锁与放行门控，不做接地电阻判级。
  作者   Author     : 道莅代码库 · PLC 编程专家（R57）
  ------------------------------------------------------------------
  边界 Boundary     :
                      一 组态闸：fAirMin > 0 且非有限拦截（R151）；
                      二 确认窗纪律：tConfirm 内持续低于下限才锁存，
                         单拍毛刺由 TON.IN 断开自然吸收；
                      三 失能即解锁：回 Idle 相、锁存清除、bPermitOk 安全侧
                         断开放行（R191 显式声明）；
                      四 锁存解除路径 = bReset 上升沿（唯一路径，R188）；
                      五 无全局变量、无外部变量声明、无物理地址寻址。
  修订记录 Revision  :
    2026-11-21  v1.0.0  R57 首版（批 4 · 序号 17）
  ==================================================================
*)

TYPE E_DL_IaiPhase :
(
    eIdle    := 0,  // 未使能：联锁停摆，放行断开 / disabled, the interlock idle, the permit open
    eRun     := 10, // 运行：风速监视 / running, the airflow watched
    eLatched := 20, // 锁存：风速欠限已确认 / latched, the underrun confirmed
    eFault   := 90  // 故障：传感失效或组态非法 / fault, a sensor failure or an illegal config
);
END_TYPE

TYPE E_DL_IaiFault :
(
    eNone       := 0, // 无成因 / no cause
    eCfgIllegal := 1, // 组态非法：下限越域（故障级，与 bError 配对）/ an illegal config
    eSensorBad  := 2, // 风速非有限（故障级，与 bError 配对）/ a non finite airflow
    eAirLow     := 3, // 风速低于下限已确认锁存（故障级，与 bError 配对）/ the underrun latched
    ePhaseBad   := 4  // 非法相位兜底（故障级，与 bError 配对）/ an illegal phase fallback
);
END_TYPE

FUNCTION_BLOCK FB_DL_IonizerAirflowInterlock
VAR_INPUT
    bEnable  : BOOL := TRUE;   // 使能，失能即解锁回空闲 [-] / enable, disabling unlocks to idle
    bReset   : BOOL := FALSE;  // 复位上升沿清锁存 [-] / reset rising edge clears the latch
    fAirflow : LREAL := 5.0;   // 风速实测 [米每秒] / the measured airflow [metre per second]
    fAirMin  : LREAL := 1.0;   // 风速下限 [米每秒]，域 大于零 / the airflow floor [metre per second], above zero
    tConfirm : TIME := T#3S;   // 欠限确认窗 [毫秒]，单拍毛刺不动作 / the confirm window [millisecond], a single glitch inert
END_VAR
VAR_OUTPUT
    bPermitOk   : BOOL := FALSE; // 放行门控出口（安全侧断开）[-] / the permit gate outlet, open on the safe side
    bIonValid   : BOOL := FALSE; // 消电离有效性出口（风速在限内）[-] / the ionization validity outlet
    bLatched    : BOOL := FALSE; // 欠限锁存电平 [-] / the underrun latch level
    tConfirmEt  : TIME := T#0S;  // 确认窗已流逝 [毫秒] / the confirm elapsed [millisecond]
    ePhase      : E_DL_IaiPhase := E_DL_IaiPhase.eIdle; // 相位出口 [枚举] / the phase outlet [enum]
    eFault      : E_DL_IaiFault := E_DL_IaiFault.eNone; // 成因出口，锁存回放 [枚举] / the cause outlet replayed
    bError      : BOOL := FALSE; // 故障锁存标志 [-] / the fault latch flag
END_VAR
VAR
    rtReset : R_TRIG; // 复位沿检测，段 0 无条件刷新 / the reset edge, refreshed unconditionally
    tonConfirm : TON; // 欠限确认窗，段 0 无条件刷新 / the confirm window, refreshed unconditionally
    _ePhase : E_DL_IaiPhase := E_DL_IaiPhase.eIdle; // 内部相位，CASE 唯一写入目标 / the internal phase
    _eFaulC : E_DL_IaiFault := E_DL_IaiFault.eNone; // 故障级成因，锁存至复位沿 / the fault cause, latched
    _bFault : BOOL := FALSE; // 故障锁存位 [-] / the fault latch bit
    _bInit  : BOOL := FALSE; // 首扫初始化完成标志（R310）/ the first scan flag
    _bInOk  : BOOL := FALSE; // 风速有限 [-] / the airflow finite
    _bCfgOk : BOOL := FALSE; // 组态域内 [-] / the config inside the domain
END_VAR

// 段 0｜定时器与沿检测无条件周期刷新（禁入分支）/ segment 0, the unconditional refresh
rtReset(CLK := bReset); // 复位沿 / the reset edge
tonConfirm(IN := (_ePhase = E_DL_IaiPhase.eRun) AND (NOT _bFault) AND _bInOk AND (fAirflow < fAirMin), PT := tConfirm); // 确认窗，IN 串运行相 / 有限 / 欠限三重闸 / the window gated by the phase, the finiteness and the underrun

// 段 1｜首扫初始化（R310）/ segment 1, the first scan
IF NOT _bInit THEN // 首扫一拍 / the first scan
    _bInit  := TRUE; // 置首扫标志 / raise the flag
    _ePhase := E_DL_IaiPhase.eRun; // 相位从运行起步（使能默认真）/ the phase starts in run
END_IF

// 段 2｜复位沿作用域：清锁存 / 迁运行相（两项逐项声明）/ segment 2, the reset edge scope
IF rtReset.Q THEN // 复位沿 / the reset edge
    _bFault := FALSE; // 作用域一：清故障锁存 / scope one, clear the fault latch
    _eFaulC := E_DL_IaiFault.eNone; // 作用域一：清成因 / scope one, clear the cause
    _ePhase := E_DL_IaiPhase.eRun; // 作用域二：迁回运行相 / scope two, back to run
END_IF

// 段 3｜组态与输入域闸（边界一）/ segment 3, the configuration and input gates
_bInOk := (fAirflow = fAirflow) AND ((fAirflow - fAirflow) = (fAirflow - fAirflow)); // 风速有限双判据 / the airflow finiteness
_bCfgOk := (fAirMin > 0.0) AND (fAirMin = fAirMin) AND ((fAirMin - fAirMin) = (fAirMin - fAirMin)) AND (tConfirm > T#0S); // 下限与确认窗域判定 / the floor and window verdict
IF (NOT _bInOk) OR (NOT _bCfgOk) THEN // 输入缺陷或组态非法 / a defect or an illegal config
    IF NOT _bFault THEN // 未锁存才迁移 / migrate only while unlatched
        _bFault := TRUE; // 置故障锁存 / raise the fault latch
        IF NOT _bInOk THEN // 传感失效优先归因（R190）/ the sensor failure first
            _eFaulC := E_DL_IaiFault.eSensorBad; // 传感成因 / the sensor cause
        ELSE // 组态非法 / the illegal config
            _eFaulC := E_DL_IaiFault.eCfgIllegal; // 组态成因 / the config cause
        END_IF
        _ePhase := E_DL_IaiPhase.eFault; // 迁故障相 / migrate to fault
    END_IF
END_IF

// 段 4｜相位机：ENUM + CASE，含 ELSE 非法相位兜底（R128）/ segment 4, the phase machine
CASE _ePhase OF

E_DL_IaiPhase.eIdle: // 未使能相 / the idle phase
    IF bEnable AND (NOT _bFault) THEN // 使能且无故障 / enabled and unfaulted
        _ePhase := E_DL_IaiPhase.eRun; // 迁运行相 / migrate to run
    END_IF

E_DL_IaiPhase.eRun: // 运行相：风速监视 / the run phase
    IF NOT bEnable THEN // 失能 / disabled
        _ePhase := E_DL_IaiPhase.eIdle; // 迁未使能相（解锁，边界三）/ migrate to idle
    ELSIF tonConfirm.Q THEN // 欠限持续确认到期（边界二）/ the underrun confirmed
        _bFault := TRUE; // 置故障锁存 / raise the fault latch
        _eFaulC := E_DL_IaiFault.eAirLow; // 故障级成因（R45 配对 bError）/ the fault cause
        _ePhase := E_DL_IaiPhase.eLatched; // 迁锁存相 / migrate to latched
    END_IF

E_DL_IaiPhase.eLatched: // 锁存相：放行断开，等复位沿或失能 / the latched phase, the permit open until the reset edge
    IF NOT bEnable THEN // 失能即解锁（边界三）/ disabling unlocks
        _bFault := FALSE; // 清故障锁存 / clear the fault latch
        _eFaulC := E_DL_IaiFault.eNone; // 清成因 / clear the cause
        _ePhase := E_DL_IaiPhase.eIdle; // 回空闲相 / back to idle
    END_IF

E_DL_IaiPhase.eFault: // 故障相：成因锁存，等复位沿或失能 / the fault phase, latched until reset or disable
    IF NOT bEnable THEN // 失能 / disabled
        _bFault := FALSE; // 清故障锁存 / clear the fault latch
        _eFaulC := E_DL_IaiFault.eNone; // 清成因 / clear the cause
        _ePhase := E_DL_IaiPhase.eIdle; // 回空闲相 / back to idle
    END_IF

ELSE // 非法相位兜底（R128）/ the illegal phase fallback
    _bFault := TRUE; // 置故障锁存 / raise the fault latch
    _eFaulC := E_DL_IaiFault.ePhaseBad; // 故障级成因（R45 配对 bError）/ the fault cause
    _ePhase := E_DL_IaiPhase.eFault; // 迁故障相 / migrate to fault
END_CASE

// 段 5｜统一出口：放行与有效性分离单点映射 / segment 5, the unified outlet
IF (_ePhase = E_DL_IaiPhase.eRun) AND (NOT _bFault) AND _bInOk AND _bCfgOk AND (fAirflow >= fAirMin) THEN // 风速在限内 / the airflow inside the band
    bPermitOk := TRUE; // 放行接通 / the permit closed
    bIonValid := TRUE; // 消电离有效 / the ionization valid
ELSE // 任何异常相放行安全侧断开（边界三）/ any abnormal phase opens the permit on the safe side
    bPermitOk := FALSE; // 放行断开 / the permit open
    bIonValid := (_ePhase = E_DL_IaiPhase.eRun) AND (NOT _bFault); // 有效性随运行相 / the validity follows the run phase
END_IF
bLatched := (_ePhase = E_DL_IaiPhase.eLatched); // 锁存电平派生 / the latch level derived
tConfirmEt := tonConfirm.ET; // 确认窗流逝出口 / the confirm elapsed outlet
ePhase := _ePhase; // 相位出口单点映射 / the phase outlet
IF _bFault THEN // 故障锁存优先 / the fault latch first
    eFault := _eFaulC; // 成因锁存回放（R152）/ the cause replayed
ELSE // 无锁存 / no latch
    eFault := E_DL_IaiFault.eNone; // 无成因 / no cause
END_IF
bError := _bFault; // 故障标志与锁存位同源 / the flag shares the latch
END_FUNCTION_BLOCK
